(* IEC 61131-3 sources: deprecated-refusr-repo/samples (part 17) *)

(* ---- 5-MUX_stows-month-choos.st ---- *)
(*
This code implements a shuffled multiplexer with 5 control bits.
The control bits are: Data[N3], Data[N24], Data[N2], Data[N10], Data[N1]
The input bits are: Data[N22], Data[N5], Data[N4], Data[N11], Data[N6], Data[N7], Data[N21], Data[N8], Data[N9], Data[N12], Data[N20], Data[N23], Data[N17], Data[N14], Data[N25], Data[N26], Data[N28], Data[N15], Data[N30], Data[N13], Data[N16], Data[N19], Data[N27], Data[N29], Data[N18], Data[N31], Data[N34], Data[N32], Data[N33], Data[N35], Data[N36], Data[N37]

The symbolic expression is:
((((((((((((((((((((((((((((((((!(((((!(IN3)) & (!(IN24))) & (!(IN2))) & (!(IN10))) & (!(IN1)))) | IN22) & ((!((((IN3 & (!(IN24))) & (!(IN2))) & (!(IN10))) & (!(IN1)))) | IN5)) & ((!(((((!(IN3)) & IN24) & (!(IN2))) & (!(IN10))) & (!(IN1)))) | IN4)) & ((!((((IN3 & IN24) & (!(IN2))) & (!(IN10))) & (!(IN1)))) | IN11)) & ((!(((((!(IN3)) & (!(IN24))) & IN2) & (!(IN10))) & (!(IN1)))) | IN6)) & ((!((((IN3 & (!(IN24))) & IN2) & (!(IN10))) & (!(IN1)))) | IN7)) & ((!(((((!(IN3)) & IN24) & IN2) & (!(IN10))) & (!(IN1)))) | IN21)) & ((!((((IN3 & IN24) & IN2) & (!(IN10))) & (!(IN1)))) | IN8)) & ((!(((((!(IN3)) & (!(IN24))) & (!(IN2))) & IN10) & (!(IN1)))) | IN9)) & ((!((((IN3 & (!(IN24))) & (!(IN2))) & IN10) & (!(IN1)))) | IN12)) & ((!(((((!(IN3)) & IN24) & (!(IN2))) & IN10) & (!(IN1)))) | IN20)) & ((!((((IN3 & IN24) & (!(IN2))) & IN10) & (!(IN1)))) | IN23)) & ((!(((((!(IN3)) & (!(IN24))) & IN2) & IN10) & (!(IN1)))) | IN17)) & ((!((((IN3 & (!(IN24))) & IN2) & IN10) & (!(IN1)))) | IN14)) & ((!(((((!(IN3)) & IN24) & IN2) & IN10) & (!(IN1)))) | IN25)) & ((!((((IN3 & IN24) & IN2) & IN10) & (!(IN1)))) | IN26)) & ((!(((((!(IN3)) & (!(IN24))) & (!(IN2))) & (!(IN10))) & IN1)) | IN28)) & ((!((((IN3 & (!(IN24))) & (!(IN2))) & (!(IN10))) & IN1)) | IN15)) & ((!(((((!(IN3)) & IN24) & (!(IN2))) & (!(IN10))) & IN1)) | IN30)) & ((!((((IN3 & IN24) & (!(IN2))) & (!(IN10))) & IN1)) | IN13)) & ((!(((((!(IN3)) & (!(IN24))) & IN2) & (!(IN10))) & IN1)) | IN16)) & ((!((((IN3 & (!(IN24))) & IN2) & (!(IN10))) & IN1)) | IN19)) & ((!(((((!(IN3)) & IN24) & IN2) & (!(IN10))) & IN1)) | IN27)) & ((!((((IN3 & IN24) & IN2) & (!(IN10))) & IN1)) | IN29)) & ((!(((((!(IN3)) & (!(IN24))) & (!(IN2))) & IN10) & IN1)) | IN18)) & ((!((((IN3 & (!(IN24))) & (!(IN2))) & IN10) & IN1)) | IN31)) & ((!(((((!(IN3)) & IN24) & (!(IN2))) & IN10) & IN1)) | IN34)) & ((!((((IN3 & IN24) & (!(IN2))) & IN10) & IN1)) | IN32)) & ((!(((((!(IN3)) & (!(IN24))) & IN2) & IN10) & IN1)) | IN33)) & ((!((((IN3 & (!(IN24))) & IN2) & IN10) & IN1)) | IN35)) & ((!(((((!(IN3)) & IN24) & IN2) & IN10) & IN1)) | IN36)) & ((!((((IN3 & IN24) & IN2) & IN10) & IN1)) | IN37)

*)

FUNCTION_BLOCK F_CollectInput
  VAR_IN_OUT
      Data : ARRAY[1..40] OF BOOL;
  END_VAR
  VAR_INPUT
      TICK  : BOOL := 0;
      IN1   : BOOL := 0;
      IN2   : BOOL := 0;
      IN3   : BOOL := 0;
      IN4   : BOOL := 0;
      IN5   : BOOL := 0;
      RESET : BOOL := FALSE;
  END_VAR
  VAR_OUTPUT
      Finished : BOOL;
  END_VAR
  VAR
      j    : USINT := 1;
      tock : BOOL  := 0;
  END_VAR
  IF NOT RESET AND tock = NOT TICK THEN
      Data[j]   := IN1;
      Data[j+1] := IN2;
      Data[j+2] := IN3;
      Data[j+3] := IN4;
      Data[j+4] := IN5;
      j := j + 5;
      tock := TICK;
  ELSE
      j := 1;
      tock := 0;
  END_IF;
  Finished := (j > 40);
END_FUNCTION_BLOCK

PROGRAM Boiler
  VAR
    Data  : ARRAY[1..40] OF BOOL;
    Ready : BOOL;
    CollectInput : F_CollectInput;
  END_VAR
  VAR
    TICK     AT %IX1.0 : BOOL;
    IN1      AT %IX0.3 : BOOL;
    IN2      AT %IX0.4 : BOOL;
    IN3      AT %IX0.5 : BOOL;
    IN4      AT %IX0.6 : BOOL;
    IN5      AT %IX0.7 : BOOL;
    OutReady AT %QX0.0 : BOOL := FALSE;
    FeedNext AT %QX0.1 : BOOL := FALSE;
    Out      AT %QX0.2 : BOOL;
  END_VAR
  CollectInput(TICK:=TICK, IN1:=IN1, IN2:=IN2, IN3:=IN3, IN4:=IN4, IN5:=IN5);
  Ready := CollectInput.Finished;
  FeedNext := 1;
  IF Ready THEN
    Out := (((((((((((((((((((((((((((((((((NOT (((((NOT Data[3]) AND (NOT Data[24])) AND (NOT Data[2])) AND (NOT Data[10])) AND (NOT Data[1]))) OR Data[22]) AND ((NOT ((((Data[3] AND (NOT Data[24])) AND (NOT Data[2])) AND (NOT Data[10])) AND (NOT Data[1]))) OR Data[5])) AND ((NOT (((((NOT Data[3]) AND Data[24]) AND (NOT Data[2])) AND (NOT Data[10])) AND (NOT Data[1]))) OR Data[4])) AND ((NOT ((((Data[3] AND Data[24]) AND (NOT Data[2])) AND (NOT Data[10])) AND (NOT Data[1]))) OR Data[11])) AND ((NOT (((((NOT Data[3]) AND (NOT Data[24])) AND Data[2]) AND (NOT Data[10])) AND (NOT Data[1]))) OR Data[6])) AND ((NOT ((((Data[3] AND (NOT Data[24])) AND Data[2]) AND (NOT Data[10])) AND (NOT Data[1]))) OR Data[7])) AND ((NOT (((((NOT Data[3]) AND Data[24]) AND Data[2]) AND (NOT Data[10])) AND (NOT Data[1]))) OR Data[21])) AND ((NOT ((((Data[3] AND Data[24]) AND Data[2]) AND (NOT Data[10])) AND (NOT Data[1]))) OR Data[8])) AND ((NOT (((((NOT Data[3]) AND (NOT Data[24])) AND (NOT Data[2])) AND Data[10]) AND (NOT Data[1]))) OR Data[9])) AND ((NOT ((((Data[3] AND (NOT Data[24])) AND (NOT Data[2])) AND Data[10]) AND (NOT Data[1]))) OR Data[12])) AND ((NOT (((((NOT Data[3]) AND Data[24]) AND (NOT Data[2])) AND Data[10]) AND (NOT Data[1]))) OR Data[20])) AND ((NOT ((((Data[3] AND Data[24]) AND (NOT Data[2])) AND Data[10]) AND (NOT Data[1]))) OR Data[23])) AND ((NOT (((((NOT Data[3]) AND (NOT Data[24])) AND Data[2]) AND Data[10]) AND (NOT Data[1]))) OR Data[17])) AND ((NOT ((((Data[3] AND (NOT Data[24])) AND Data[2]) AND Data[10]) AND (NOT Data[1]))) OR Data[14])) AND ((NOT (((((NOT Data[3]) AND Data[24]) AND Data[2]) AND Data[10]) AND (NOT Data[1]))) OR Data[25])) AND ((NOT ((((Data[3] AND Data[24]) AND Data[2]) AND Data[10]) AND (NOT Data[1]))) OR Data[26])) AND ((NOT (((((NOT Data[3]) AND (NOT Data[24])) AND (NOT Data[2])) AND (NOT Data[10])) AND Data[1])) OR Data[28])) AND ((NOT ((((Data[3] AND (NOT Data[24])) AND (NOT Data[2])) AND (NOT Data[10])) AND Data[1])) OR Data[15])) AND ((NOT (((((NOT Data[3]) AND Data[24]) AND (NOT Data[2])) AND (NOT Data[10])) AND Data[1])) OR Data[30])) AND ((NOT ((((Data[3] AND Data[24]) AND (NOT Data[2])) AND (NOT Data[10])) AND Data[1])) OR Data[13])) AND ((NOT (((((NOT Data[3]) AND (NOT Data[24])) AND Data[2]) AND (NOT Data[10])) AND Data[1])) OR Data[16])) AND ((NOT ((((Data[3] AND (NOT Data[24])) AND Data[2]) AND (NOT Data[10])) AND Data[1])) OR Data[19])) AND ((NOT (((((NOT Data[3]) AND Data[24]) AND Data[2]) AND (NOT Data[10])) AND Data[1])) OR Data[27])) AND ((NOT ((((Data[3] AND Data[24]) AND Data[2]) AND (NOT Data[10])) AND Data[1])) OR Data[29])) AND ((NOT (((((NOT Data[3]) AND (NOT Data[24])) AND (NOT Data[2])) AND Data[10]) AND Data[1])) OR Data[18])) AND ((NOT ((((Data[3] AND (NOT Data[24])) AND (NOT Data[2])) AND Data[10]) AND Data[1])) OR Data[31])) AND ((NOT (((((NOT Data[3]) AND Data[24]) AND (NOT Data[2])) AND Data[10]) AND Data[1])) OR Data[34])) AND ((NOT ((((Data[3] AND Data[24]) AND (NOT Data[2])) AND Data[10]) AND Data[1])) OR Data[32])) AND ((NOT (((((NOT Data[3]) AND (NOT Data[24])) AND Data[2]) AND Data[10]) AND Data[1])) OR Data[33])) AND ((NOT ((((Data[3] AND (NOT Data[24])) AND Data[2]) AND Data[10]) AND Data[1])) OR Data[35])) AND ((NOT (((((NOT Data[3]) AND Data[24]) AND Data[2]) AND Data[10]) AND Data[1])) OR Data[36])) AND ((NOT ((((Data[3] AND Data[24]) AND Data[2]) AND Data[10]) AND Data[1])) OR Data[37]));
    OutReady := 1;
    CollectInput(RESET:=TRUE);
  END_IF;
END_PROGRAM

CONFIGURATION Config0
  RESOURCE Res0 ON PLC
    TASK task0(INTERVAL := T#20ms,PRIORITY := 0);
    PROGRAM instance0 WITH task0 : Boiler;
  END_RESOURCE
END_CONFIGURATION

(* ---- 5-MUX_strop-getup-abyss.st ---- *)
(*
This code implements a shuffled multiplexer with 5 control bits.
The control bits are: Data[N2], Data[N8], Data[N3], Data[N22], Data[N21]
The input bits are: Data[N20], Data[N25], Data[N5], Data[N1], Data[N6], Data[N24], Data[N23], Data[N26], Data[N27], Data[N7], Data[N28], Data[N29], Data[N10], Data[N30], Data[N33], Data[N9], Data[N4], Data[N11], Data[N12], Data[N31], Data[N32], Data[N36], Data[N34], Data[N37], Data[N15], Data[N35], Data[N14], Data[N13], Data[N17], Data[N18], Data[N16], Data[N19]

The symbolic expression is:
((((((((((((((((((((((((((((((((!(((((!(IN2)) & (!(IN8))) & (!(IN3))) & (!(IN22))) & (!(IN21)))) | IN20) & ((!((((IN2 & (!(IN8))) & (!(IN3))) & (!(IN22))) & (!(IN21)))) | IN25)) & ((!(((((!(IN2)) & IN8) & (!(IN3))) & (!(IN22))) & (!(IN21)))) | IN5)) & ((!((((IN2 & IN8) & (!(IN3))) & (!(IN22))) & (!(IN21)))) | IN1)) & ((!(((((!(IN2)) & (!(IN8))) & IN3) & (!(IN22))) & (!(IN21)))) | IN6)) & ((!((((IN2 & (!(IN8))) & IN3) & (!(IN22))) & (!(IN21)))) | IN24)) & ((!(((((!(IN2)) & IN8) & IN3) & (!(IN22))) & (!(IN21)))) | IN23)) & ((!((((IN2 & IN8) & IN3) & (!(IN22))) & (!(IN21)))) | IN26)) & ((!(((((!(IN2)) & (!(IN8))) & (!(IN3))) & IN22) & (!(IN21)))) | IN27)) & ((!((((IN2 & (!(IN8))) & (!(IN3))) & IN22) & (!(IN21)))) | IN7)) & ((!(((((!(IN2)) & IN8) & (!(IN3))) & IN22) & (!(IN21)))) | IN28)) & ((!((((IN2 & IN8) & (!(IN3))) & IN22) & (!(IN21)))) | IN29)) & ((!(((((!(IN2)) & (!(IN8))) & IN3) & IN22) & (!(IN21)))) | IN10)) & ((!((((IN2 & (!(IN8))) & IN3) & IN22) & (!(IN21)))) | IN30)) & ((!(((((!(IN2)) & IN8) & IN3) & IN22) & (!(IN21)))) | IN33)) & ((!((((IN2 & IN8) & IN3) & IN22) & (!(IN21)))) | IN9)) & ((!(((((!(IN2)) & (!(IN8))) & (!(IN3))) & (!(IN22))) & IN21)) | IN4)) & ((!((((IN2 & (!(IN8))) & (!(IN3))) & (!(IN22))) & IN21)) | IN11)) & ((!(((((!(IN2)) & IN8) & (!(IN3))) & (!(IN22))) & IN21)) | IN12)) & ((!((((IN2 & IN8) & (!(IN3))) & (!(IN22))) & IN21)) | IN31)) & ((!(((((!(IN2)) & (!(IN8))) & IN3) & (!(IN22))) & IN21)) | IN32)) & ((!((((IN2 & (!(IN8))) & IN3) & (!(IN22))) & IN21)) | IN36)) & ((!(((((!(IN2)) & IN8) & IN3) & (!(IN22))) & IN21)) | IN34)) & ((!((((IN2 & IN8) & IN3) & (!(IN22))) & IN21)) | IN37)) & ((!(((((!(IN2)) & (!(IN8))) & (!(IN3))) & IN22) & IN21)) | IN15)) & ((!((((IN2 & (!(IN8))) & (!(IN3))) & IN22) & IN21)) | IN35)) & ((!(((((!(IN2)) & IN8) & (!(IN3))) & IN22) & IN21)) | IN14)) & ((!((((IN2 & IN8) & (!(IN3))) & IN22) & IN21)) | IN13)) & ((!(((((!(IN2)) & (!(IN8))) & IN3) & IN22) & IN21)) | IN17)) & ((!((((IN2 & (!(IN8))) & IN3) & IN22) & IN21)) | IN18)) & ((!(((((!(IN2)) & IN8) & IN3) & IN22) & IN21)) | IN16)) & ((!((((IN2 & IN8) & IN3) & IN22) & IN21)) | IN19)

*)

FUNCTION_BLOCK F_CollectInput
  VAR_IN_OUT
      Data : ARRAY[1..40] OF BOOL;
  END_VAR
  VAR_INPUT
      TICK  : BOOL := 0;
      IN1   : BOOL := 0;
      IN2   : BOOL := 0;
      IN3   : BOOL := 0;
      IN4   : BOOL := 0;
      IN5   : BOOL := 0;
      RESET : BOOL := FALSE;
  END_VAR
  VAR_OUTPUT
      Finished : BOOL;
  END_VAR
  VAR
      j    : USINT := 1;
      tock : BOOL  := 0;
  END_VAR
  IF NOT RESET AND tock = NOT TICK THEN
      Data[j]   := IN1;
      Data[j+1] := IN2;
      Data[j+2] := IN3;
      Data[j+3] := IN4;
      Data[j+4] := IN5;
      j := j + 5;
      tock := TICK;
  ELSE
      j := 1;
      tock := 0;
  END_IF;
  Finished := (j > 40);
END_FUNCTION_BLOCK

PROGRAM Boiler
  VAR
    Data  : ARRAY[1..40] OF BOOL;
    Ready : BOOL;
    CollectInput : F_CollectInput;
  END_VAR
  VAR
    TICK     AT %IX1.0 : BOOL;
    IN1      AT %IX0.3 : BOOL;
    IN2      AT %IX0.4 : BOOL;
    IN3      AT %IX0.5 : BOOL;
    IN4      AT %IX0.6 : BOOL;
    IN5      AT %IX0.7 : BOOL;
    OutReady AT %QX0.0 : BOOL := FALSE;
    FeedNext AT %QX0.1 : BOOL := FALSE;
    Out      AT %QX0.2 : BOOL;
  END_VAR
  CollectInput(TICK:=TICK, IN1:=IN1, IN2:=IN2, IN3:=IN3, IN4:=IN4, IN5:=IN5);
  Ready := CollectInput.Finished;
  FeedNext := 1;
  IF Ready THEN
    Out := (((((((((((((((((((((((((((((((((NOT (((((NOT Data[2]) AND (NOT Data[8])) AND (NOT Data[3])) AND (NOT Data[22])) AND (NOT Data[21]))) OR Data[20]) AND ((NOT ((((Data[2] AND (NOT Data[8])) AND (NOT Data[3])) AND (NOT Data[22])) AND (NOT Data[21]))) OR Data[25])) AND ((NOT (((((NOT Data[2]) AND Data[8]) AND (NOT Data[3])) AND (NOT Data[22])) AND (NOT Data[21]))) OR Data[5])) AND ((NOT ((((Data[2] AND Data[8]) AND (NOT Data[3])) AND (NOT Data[22])) AND (NOT Data[21]))) OR Data[1])) AND ((NOT (((((NOT Data[2]) AND (NOT Data[8])) AND Data[3]) AND (NOT Data[22])) AND (NOT Data[21]))) OR Data[6])) AND ((NOT ((((Data[2] AND (NOT Data[8])) AND Data[3]) AND (NOT Data[22])) AND (NOT Data[21]))) OR Data[24])) AND ((NOT (((((NOT Data[2]) AND Data[8]) AND Data[3]) AND (NOT Data[22])) AND (NOT Data[21]))) OR Data[23])) AND ((NOT ((((Data[2] AND Data[8]) AND Data[3]) AND (NOT Data[22])) AND (NOT Data[21]))) OR Data[26])) AND ((NOT (((((NOT Data[2]) AND (NOT Data[8])) AND (NOT Data[3])) AND Data[22]) AND (NOT Data[21]))) OR Data[27])) AND ((NOT ((((Data[2] AND (NOT Data[8])) AND (NOT Data[3])) AND Data[22]) AND (NOT Data[21]))) OR Data[7])) AND ((NOT (((((NOT Data[2]) AND Data[8]) AND (NOT Data[3])) AND Data[22]) AND (NOT Data[21]))) OR Data[28])) AND ((NOT ((((Data[2] AND Data[8]) AND (NOT Data[3])) AND Data[22]) AND (NOT Data[21]))) OR Data[29])) AND ((NOT (((((NOT Data[2]) AND (NOT Data[8])) AND Data[3]) AND Data[22]) AND (NOT Data[21]))) OR Data[10])) AND ((NOT ((((Data[2] AND (NOT Data[8])) AND Data[3]) AND Data[22]) AND (NOT Data[21]))) OR Data[30])) AND ((NOT (((((NOT Data[2]) AND Data[8]) AND Data[3]) AND Data[22]) AND (NOT Data[21]))) OR Data[33])) AND ((NOT ((((Data[2] AND Data[8]) AND Data[3]) AND Data[22]) AND (NOT Data[21]))) OR Data[9])) AND ((NOT (((((NOT Data[2]) AND (NOT Data[8])) AND (NOT Data[3])) AND (NOT Data[22])) AND Data[21])) OR Data[4])) AND ((NOT ((((Data[2] AND (NOT Data[8])) AND (NOT Data[3])) AND (NOT Data[22])) AND Data[21])) OR Data[11])) AND ((NOT (((((NOT Data[2]) AND Data[8]) AND (NOT Data[3])) AND (NOT Data[22])) AND Data[21])) OR Data[12])) AND ((NOT ((((Data[2] AND Data[8]) AND (NOT Data[3])) AND (NOT Data[22])) AND Data[21])) OR Data[31])) AND ((NOT (((((NOT Data[2]) AND (NOT Data[8])) AND Data[3]) AND (NOT Data[22])) AND Data[21])) OR Data[32])) AND ((NOT ((((Data[2] AND (NOT Data[8])) AND Data[3]) AND (NOT Data[22])) AND Data[21])) OR Data[36])) AND ((NOT (((((NOT Data[2]) AND Data[8]) AND Data[3]) AND (NOT Data[22])) AND Data[21])) OR Data[34])) AND ((NOT ((((Data[2] AND Data[8]) AND Data[3]) AND (NOT Data[22])) AND Data[21])) OR Data[37])) AND ((NOT (((((NOT Data[2]) AND (NOT Data[8])) AND (NOT Data[3])) AND Data[22]) AND Data[21])) OR Data[15])) AND ((NOT ((((Data[2] AND (NOT Data[8])) AND (NOT Data[3])) AND Data[22]) AND Data[21])) OR Data[35])) AND ((NOT (((((NOT Data[2]) AND Data[8]) AND (NOT Data[3])) AND Data[22]) AND Data[21])) OR Data[14])) AND ((NOT ((((Data[2] AND Data[8]) AND (NOT Data[3])) AND Data[22]) AND Data[21])) OR Data[13])) AND ((NOT (((((NOT Data[2]) AND (NOT Data[8])) AND Data[3]) AND Data[22]) AND Data[21])) OR Data[17])) AND ((NOT ((((Data[2] AND (NOT Data[8])) AND Data[3]) AND Data[22]) AND Data[21])) OR Data[18])) AND ((NOT (((((NOT Data[2]) AND Data[8]) AND Data[3]) AND Data[22]) AND Data[21])) OR Data[16])) AND ((NOT ((((Data[2] AND Data[8]) AND Data[3]) AND Data[22]) AND Data[21])) OR Data[19]));
    OutReady := 1;
    CollectInput(RESET:=TRUE);
  END_IF;
END_PROGRAM

CONFIGURATION Config0
  RESOURCE Res0 ON PLC
    TASK task0(INTERVAL := T#20ms,PRIORITY := 0);
    PROGRAM instance0 WITH task0 : Boiler;
  END_RESOURCE
END_CONFIGURATION

(* ---- 5-MUX_supes-buret-rules.st ---- *)
(*
This code implements a shuffled multiplexer with 5 control bits.
The control bits are: Data[N20], Data[N2], Data[N3], Data[N1], Data[N4]
The input bits are: Data[N7], Data[N21], Data[N22], Data[N25], Data[N5], Data[N24], Data[N9], Data[N10], Data[N8], Data[N26], Data[N23], Data[N6], Data[N11], Data[N12], Data[N28], Data[N13], Data[N14], Data[N30], Data[N15], Data[N29], Data[N16], Data[N17], Data[N18], Data[N19], Data[N27], Data[N31], Data[N33], Data[N35], Data[N32], Data[N34], Data[N37], Data[N36]

The symbolic expression is:
((((((((((((((((((((((((((((((((!(((((!(IN20)) & (!(IN2))) & (!(IN3))) & (!(IN1))) & (!(IN4)))) | IN7) & ((!((((IN20 & (!(IN2))) & (!(IN3))) & (!(IN1))) & (!(IN4)))) | IN21)) & ((!(((((!(IN20)) & IN2) & (!(IN3))) & (!(IN1))) & (!(IN4)))) | IN22)) & ((!((((IN20 & IN2) & (!(IN3))) & (!(IN1))) & (!(IN4)))) | IN25)) & ((!(((((!(IN20)) & (!(IN2))) & IN3) & (!(IN1))) & (!(IN4)))) | IN5)) & ((!((((IN20 & (!(IN2))) & IN3) & (!(IN1))) & (!(IN4)))) | IN24)) & ((!(((((!(IN20)) & IN2) & IN3) & (!(IN1))) & (!(IN4)))) | IN9)) & ((!((((IN20 & IN2) & IN3) & (!(IN1))) & (!(IN4)))) | IN10)) & ((!(((((!(IN20)) & (!(IN2))) & (!(IN3))) & IN1) & (!(IN4)))) | IN8)) & ((!((((IN20 & (!(IN2))) & (!(IN3))) & IN1) & (!(IN4)))) | IN26)) & ((!(((((!(IN20)) & IN2) & (!(IN3))) & IN1) & (!(IN4)))) | IN23)) & ((!((((IN20 & IN2) & (!(IN3))) & IN1) & (!(IN4)))) | IN6)) & ((!(((((!(IN20)) & (!(IN2))) & IN3) & IN1) & (!(IN4)))) | IN11)) & ((!((((IN20 & (!(IN2))) & IN3) & IN1) & (!(IN4)))) | IN12)) & ((!(((((!(IN20)) & IN2) & IN3) & IN1) & (!(IN4)))) | IN28)) & ((!((((IN20 & IN2) & IN3) & IN1) & (!(IN4)))) | IN13)) & ((!(((((!(IN20)) & (!(IN2))) & (!(IN3))) & (!(IN1))) & IN4)) | IN14)) & ((!((((IN20 & (!(IN2))) & (!(IN3))) & (!(IN1))) & IN4)) | IN30)) & ((!(((((!(IN20)) & IN2) & (!(IN3))) & (!(IN1))) & IN4)) | IN15)) & ((!((((IN20 & IN2) & (!(IN3))) & (!(IN1))) & IN4)) | IN29)) & ((!(((((!(IN20)) & (!(IN2))) & IN3) & (!(IN1))) & IN4)) | IN16)) & ((!((((IN20 & (!(IN2))) & IN3) & (!(IN1))) & IN4)) | IN17)) & ((!(((((!(IN20)) & IN2) & IN3) & (!(IN1))) & IN4)) | IN18)) & ((!((((IN20 & IN2) & IN3) & (!(IN1))) & IN4)) | IN19)) & ((!(((((!(IN20)) & (!(IN2))) & (!(IN3))) & IN1) & IN4)) | IN27)) & ((!((((IN20 & (!(IN2))) & (!(IN3))) & IN1) & IN4)) | IN31)) & ((!(((((!(IN20)) & IN2) & (!(IN3))) & IN1) & IN4)) | IN33)) & ((!((((IN20 & IN2) & (!(IN3))) & IN1) & IN4)) | IN35)) & ((!(((((!(IN20)) & (!(IN2))) & IN3) & IN1) & IN4)) | IN32)) & ((!((((IN20 & (!(IN2))) & IN3) & IN1) & IN4)) | IN34)) & ((!(((((!(IN20)) & IN2) & IN3) & IN1) & IN4)) | IN37)) & ((!((((IN20 & IN2) & IN3) & IN1) & IN4)) | IN36)

*)

FUNCTION_BLOCK F_CollectInput
  VAR_IN_OUT
      Data : ARRAY[1..40] OF BOOL;
  END_VAR
  VAR_INPUT
      TICK  : BOOL := 0;
      IN1   : BOOL := 0;
      IN2   : BOOL := 0;
      IN3   : BOOL := 0;
      IN4   : BOOL := 0;
      IN5   : BOOL := 0;
      RESET : BOOL := FALSE;
  END_VAR
  VAR_OUTPUT
      Finished : BOOL;
  END_VAR
  VAR
      j    : USINT := 1;
      tock : BOOL  := 0;
  END_VAR
  IF NOT RESET AND tock = NOT TICK THEN
      Data[j]   := IN1;
      Data[j+1] := IN2;
      Data[j+2] := IN3;
      Data[j+3] := IN4;
      Data[j+4] := IN5;
      j := j + 5;
      tock := TICK;
  ELSE
      j := 1;
      tock := 0;
  END_IF;
  Finished := (j > 40);
END_FUNCTION_BLOCK

PROGRAM Boiler
  VAR
    Data  : ARRAY[1..40] OF BOOL;
    Ready : BOOL;
    CollectInput : F_CollectInput;
  END_VAR
  VAR
    TICK     AT %IX1.0 : BOOL;
    IN1      AT %IX0.3 : BOOL;
    IN2      AT %IX0.4 : BOOL;
    IN3      AT %IX0.5 : BOOL;
    IN4      AT %IX0.6 : BOOL;
    IN5      AT %IX0.7 : BOOL;
    OutReady AT %QX0.0 : BOOL := FALSE;
    FeedNext AT %QX0.1 : BOOL := FALSE;
    Out      AT %QX0.2 : BOOL;
  END_VAR
  CollectInput(TICK:=TICK, IN1:=IN1, IN2:=IN2, IN3:=IN3, IN4:=IN4, IN5:=IN5);
  Ready := CollectInput.Finished;
  FeedNext := 1;
  IF Ready THEN
    Out := (((((((((((((((((((((((((((((((((NOT (((((NOT Data[20]) AND (NOT Data[2])) AND (NOT Data[3])) AND (NOT Data[1])) AND (NOT Data[4]))) OR Data[7]) AND ((NOT ((((Data[20] AND (NOT Data[2])) AND (NOT Data[3])) AND (NOT Data[1])) AND (NOT Data[4]))) OR Data[21])) AND ((NOT (((((NOT Data[20]) AND Data[2]) AND (NOT Data[3])) AND (NOT Data[1])) AND (NOT Data[4]))) OR Data[22])) AND ((NOT ((((Data[20] AND Data[2]) AND (NOT Data[3])) AND (NOT Data[1])) AND (NOT Data[4]))) OR Data[25])) AND ((NOT (((((NOT Data[20]) AND (NOT Data[2])) AND Data[3]) AND (NOT Data[1])) AND (NOT Data[4]))) OR Data[5])) AND ((NOT ((((Data[20] AND (NOT Data[2])) AND Data[3]) AND (NOT Data[1])) AND (NOT Data[4]))) OR Data[24])) AND ((NOT (((((NOT Data[20]) AND Data[2]) AND Data[3]) AND (NOT Data[1])) AND (NOT Data[4]))) OR Data[9])) AND ((NOT ((((Data[20] AND Data[2]) AND Data[3]) AND (NOT Data[1])) AND (NOT Data[4]))) OR Data[10])) AND ((NOT (((((NOT Data[20]) AND (NOT Data[2])) AND (NOT Data[3])) AND Data[1]) AND (NOT Data[4]))) OR Data[8])) AND ((NOT ((((Data[20] AND (NOT Data[2])) AND (NOT Data[3])) AND Data[1]) AND (NOT Data[4]))) OR Data[26])) AND ((NOT (((((NOT Data[20]) AND Data[2]) AND (NOT Data[3])) AND Data[1]) AND (NOT Data[4]))) OR Data[23])) AND ((NOT ((((Data[20] AND Data[2]) AND (NOT Data[3])) AND Data[1]) AND (NOT Data[4]))) OR Data[6])) AND ((NOT (((((NOT Data[20]) AND (NOT Data[2])) AND Data[3]) AND Data[1]) AND (NOT Data[4]))) OR Data[11])) AND ((NOT ((((Data[20] AND (NOT Data[2])) AND Data[3]) AND Data[1]) AND (NOT Data[4]))) OR Data[12])) AND ((NOT (((((NOT Data[20]) AND Data[2]) AND Data[3]) AND Data[1]) AND (NOT Data[4]))) OR Data[28])) AND ((NOT ((((Data[20] AND Data[2]) AND Data[3]) AND Data[1]) AND (NOT Data[4]))) OR Data[13])) AND ((NOT (((((NOT Data[20]) AND (NOT Data[2])) AND (NOT Data[3])) AND (NOT Data[1])) AND Data[4])) OR Data[14])) AND ((NOT ((((Data[20] AND (NOT Data[2])) AND (NOT Data[3])) AND (NOT Data[1])) AND Data[4])) OR Data[30])) AND ((NOT (((((NOT Data[20]) AND Data[2]) AND (NOT Data[3])) AND (NOT Data[1])) AND Data[4])) OR Data[15])) AND ((NOT ((((Data[20] AND Data[2]) AND (NOT Data[3])) AND (NOT Data[1])) AND Data[4])) OR Data[29])) AND ((NOT (((((NOT Data[20]) AND (NOT Data[2])) AND Data[3]) AND (NOT Data[1])) AND Data[4])) OR Data[16])) AND ((NOT ((((Data[20] AND (NOT Data[2])) AND Data[3]) AND (NOT Data[1])) AND Data[4])) OR Data[17])) AND ((NOT (((((NOT Data[20]) AND Data[2]) AND Data[3]) AND (NOT Data[1])) AND Data[4])) OR Data[18])) AND ((NOT ((((Data[20] AND Data[2]) AND Data[3]) AND (NOT Data[1])) AND Data[4])) OR Data[19])) AND ((NOT (((((NOT Data[20]) AND (NOT Data[2])) AND (NOT Data[3])) AND Data[1]) AND Data[4])) OR Data[27])) AND ((NOT ((((Data[20] AND (NOT Data[2])) AND (NOT Data[3])) AND Data[1]) AND Data[4])) OR Data[31])) AND ((NOT (((((NOT Data[20]) AND Data[2]) AND (NOT Data[3])) AND Data[1]) AND Data[4])) OR Data[33])) AND ((NOT ((((Data[20] AND Data[2]) AND (NOT Data[3])) AND Data[1]) AND Data[4])) OR Data[35])) AND ((NOT (((((NOT Data[20]) AND (NOT Data[2])) AND Data[3]) AND Data[1]) AND Data[4])) OR Data[32])) AND ((NOT ((((Data[20] AND (NOT Data[2])) AND Data[3]) AND Data[1]) AND Data[4])) OR Data[34])) AND ((NOT (((((NOT Data[20]) AND Data[2]) AND Data[3]) AND Data[1]) AND Data[4])) OR Data[37])) AND ((NOT ((((Data[20] AND Data[2]) AND Data[3]) AND Data[1]) AND Data[4])) OR Data[36]));
    OutReady := 1;
    CollectInput(RESET:=TRUE);
  END_IF;
END_PROGRAM

CONFIGURATION Config0
  RESOURCE Res0 ON PLC
    TASK task0(INTERVAL := T#20ms,PRIORITY := 0);
    PROGRAM instance0 WITH task0 : Boiler;
  END_RESOURCE
END_CONFIGURATION

(* ---- 5-MUX_swart-booty-dozes.st ---- *)
(*
This code implements a shuffled multiplexer with 5 control bits.
The control bits are: Data[N20], Data[N21], Data[N2], Data[N1], Data[N3]
The input bits are: Data[N22], Data[N27], Data[N6], Data[N5], Data[N4], Data[N23], Data[N29], Data[N24], Data[N25], Data[N30], Data[N28], Data[N7], Data[N9], Data[N8], Data[N10], Data[N26], Data[N11], Data[N12], Data[N14], Data[N13], Data[N34], Data[N31], Data[N15], Data[N17], Data[N18], Data[N19], Data[N33], Data[N16], Data[N35], Data[N32], Data[N36], Data[N37]

The symbolic expression is:
((((((((((((((((((((((((((((((((!(((((!(IN20)) & (!(IN21))) & (!(IN2))) & (!(IN1))) & (!(IN3)))) | IN22) & ((!((((IN20 & (!(IN21))) & (!(IN2))) & (!(IN1))) & (!(IN3)))) | IN27)) & ((!(((((!(IN20)) & IN21) & (!(IN2))) & (!(IN1))) & (!(IN3)))) | IN6)) & ((!((((IN20 & IN21) & (!(IN2))) & (!(IN1))) & (!(IN3)))) | IN5)) & ((!(((((!(IN20)) & (!(IN21))) & IN2) & (!(IN1))) & (!(IN3)))) | IN4)) & ((!((((IN20 & (!(IN21))) & IN2) & (!(IN1))) & (!(IN3)))) | IN23)) & ((!(((((!(IN20)) & IN21) & IN2) & (!(IN1))) & (!(IN3)))) | IN29)) & ((!((((IN20 & IN21) & IN2) & (!(IN1))) & (!(IN3)))) | IN24)) & ((!(((((!(IN20)) & (!(IN21))) & (!(IN2))) & IN1) & (!(IN3)))) | IN25)) & ((!((((IN20 & (!(IN21))) & (!(IN2))) & IN1) & (!(IN3)))) | IN30)) & ((!(((((!(IN20)) & IN21) & (!(IN2))) & IN1) & (!(IN3)))) | IN28)) & ((!((((IN20 & IN21) & (!(IN2))) & IN1) & (!(IN3)))) | IN7)) & ((!(((((!(IN20)) & (!(IN21))) & IN2) & IN1) & (!(IN3)))) | IN9)) & ((!((((IN20 & (!(IN21))) & IN2) & IN1) & (!(IN3)))) | IN8)) & ((!(((((!(IN20)) & IN21) & IN2) & IN1) & (!(IN3)))) | IN10)) & ((!((((IN20 & IN21) & IN2) & IN1) & (!(IN3)))) | IN26)) & ((!(((((!(IN20)) & (!(IN21))) & (!(IN2))) & (!(IN1))) & IN3)) | IN11)) & ((!((((IN20 & (!(IN21))) & (!(IN2))) & (!(IN1))) & IN3)) | IN12)) & ((!(((((!(IN20)) & IN21) & (!(IN2))) & (!(IN1))) & IN3)) | IN14)) & ((!((((IN20 & IN21) & (!(IN2))) & (!(IN1))) & IN3)) | IN13)) & ((!(((((!(IN20)) & (!(IN21))) & IN2) & (!(IN1))) & IN3)) | IN34)) & ((!((((IN20 & (!(IN21))) & IN2) & (!(IN1))) & IN3)) | IN31)) & ((!(((((!(IN20)) & IN21) & IN2) & (!(IN1))) & IN3)) | IN15)) & ((!((((IN20 & IN21) & IN2) & (!(IN1))) & IN3)) | IN17)) & ((!(((((!(IN20)) & (!(IN21))) & (!(IN2))) & IN1) & IN3)) | IN18)) & ((!((((IN20 & (!(IN21))) & (!(IN2))) & IN1) & IN3)) | IN19)) & ((!(((((!(IN20)) & IN21) & (!(IN2))) & IN1) & IN3)) | IN33)) & ((!((((IN20 & IN21) & (!(IN2))) & IN1) & IN3)) | IN16)) & ((!(((((!(IN20)) & (!(IN21))) & IN2) & IN1) & IN3)) | IN35)) & ((!((((IN20 & (!(IN21))) & IN2) & IN1) & IN3)) | IN32)) & ((!(((((!(IN20)) & IN21) & IN2) & IN1) & IN3)) | IN36)) & ((!((((IN20 & IN21) & IN2) & IN1) & IN3)) | IN37)

*)

FUNCTION_BLOCK F_CollectInput
  VAR_IN_OUT
      Data : ARRAY[1..40] OF BOOL;
  END_VAR
  VAR_INPUT
      TICK  : BOOL := 0;
      IN1   : BOOL := 0;
      IN2   : BOOL := 0;
      IN3   : BOOL := 0;
      IN4   : BOOL := 0;
      IN5   : BOOL := 0;
      RESET : BOOL := FALSE;
  END_VAR
  VAR_OUTPUT
      Finished : BOOL;
  END_VAR
  VAR
      j    : USINT := 1;
      tock : BOOL  := 0;
  END_VAR
  IF NOT RESET AND tock = NOT TICK THEN
      Data[j]   := IN1;
      Data[j+1] := IN2;
      Data[j+2] := IN3;
      Data[j+3] := IN4;
      Data[j+4] := IN5;
      j := j + 5;
      tock := TICK;
  ELSE
      j := 1;
      tock := 0;
  END_IF;
  Finished := (j > 40);
END_FUNCTION_BLOCK

PROGRAM Boiler
  VAR
    Data  : ARRAY[1..40] OF BOOL;
    Ready : BOOL;
    CollectInput : F_CollectInput;
  END_VAR
  VAR
    TICK     AT %IX1.0 : BOOL;
    IN1      AT %IX0.3 : BOOL;
    IN2      AT %IX0.4 : BOOL;
    IN3      AT %IX0.5 : BOOL;
    IN4      AT %IX0.6 : BOOL;
    IN5      AT %IX0.7 : BOOL;
    OutReady AT %QX0.0 : BOOL := FALSE;
    FeedNext AT %QX0.1 : BOOL := FALSE;
    Out      AT %QX0.2 : BOOL;
  END_VAR
  CollectInput(TICK:=TICK, IN1:=IN1, IN2:=IN2, IN3:=IN3, IN4:=IN4, IN5:=IN5);
  Ready := CollectInput.Finished;
  FeedNext := 1;
  IF Ready THEN
    Out := (((((((((((((((((((((((((((((((((NOT (((((NOT Data[20]) AND (NOT Data[21])) AND (NOT Data[2])) AND (NOT Data[1])) AND (NOT Data[3]))) OR Data[22]) AND ((NOT ((((Data[20] AND (NOT Data[21])) AND (NOT Data[2])) AND (NOT Data[1])) AND (NOT Data[3]))) OR Data[27])) AND ((NOT (((((NOT Data[20]) AND Data[21]) AND (NOT Data[2])) AND (NOT Data[1])) AND (NOT Data[3]))) OR Data[6])) AND ((NOT ((((Data[20] AND Data[21]) AND (NOT Data[2])) AND (NOT Data[1])) AND (NOT Data[3]))) OR Data[5])) AND ((NOT (((((NOT Data[20]) AND (NOT Data[21])) AND Data[2]) AND (NOT Data[1])) AND (NOT Data[3]))) OR Data[4])) AND ((NOT ((((Data[20] AND (NOT Data[21])) AND Data[2]) AND (NOT Data[1])) AND (NOT Data[3]))) OR Data[23])) AND ((NOT (((((NOT Data[20]) AND Data[21]) AND Data[2]) AND (NOT Data[1])) AND (NOT Data[3]))) OR Data[29])) AND ((NOT ((((Data[20] AND Data[21]) AND Data[2]) AND (NOT Data[1])) AND (NOT Data[3]))) OR Data[24])) AND ((NOT (((((NOT Data[20]) AND (NOT Data[21])) AND (NOT Data[2])) AND Data[1]) AND (NOT Data[3]))) OR Data[25])) AND ((NOT ((((Data[20] AND (NOT Data[21])) AND (NOT Data[2])) AND Data[1]) AND (NOT Data[3]))) OR Data[30])) AND ((NOT (((((NOT Data[20]) AND Data[21]) AND (NOT Data[2])) AND Data[1]) AND (NOT Data[3]))) OR Data[28])) AND ((NOT ((((Data[20] AND Data[21]) AND (NOT Data[2])) AND Data[1]) AND (NOT Data[3]))) OR Data[7])) AND ((NOT (((((NOT Data[20]) AND (NOT Data[21])) AND Data[2]) AND Data[1]) AND (NOT Data[3]))) OR Data[9])) AND ((NOT ((((Data[20] AND (NOT Data[21])) AND Data[2]) AND Data[1]) AND (NOT Data[3]))) OR Data[8])) AND ((NOT (((((NOT Data[20]) AND Data[21]) AND Data[2]) AND Data[1]) AND (NOT Data[3]))) OR Data[10])) AND ((NOT ((((Data[20] AND Data[21]) AND Data[2]) AND Data[1]) AND (NOT Data[3]))) OR Data[26])) AND ((NOT (((((NOT Data[20]) AND (NOT Data[21])) AND (NOT Data[2])) AND (NOT Data[1])) AND Data[3])) OR Data[11])) AND ((NOT ((((Data[20] AND (NOT Data[21])) AND (NOT Data[2])) AND (NOT Data[1])) AND Data[3])) OR Data[12])) AND ((NOT (((((NOT Data[20]) AND Data[21]) AND (NOT Data[2])) AND (NOT Data[1])) AND Data[3])) OR Data[14])) AND ((NOT ((((Data[20] AND Data[21]) AND (NOT Data[2])) AND (NOT Data[1])) AND Data[3])) OR Data[13])) AND ((NOT (((((NOT Data[20]) AND (NOT Data[21])) AND Data[2]) AND (NOT Data[1])) AND Data[3])) OR Data[34])) AND ((NOT ((((Data[20] AND (NOT Data[21])) AND Data[2]) AND (NOT Data[1])) AND Data[3])) OR Data[31])) AND ((NOT (((((NOT Data[20]) AND Data[21]) AND Data[2]) AND (NOT Data[1])) AND Data[3])) OR Data[15])) AND ((NOT ((((Data[20] AND Data[21]) AND Data[2]) AND (NOT Data[1])) AND Data[3])) OR Data[17])) AND ((NOT (((((NOT Data[20]) AND (NOT Data[21])) AND (NOT Data[2])) AND Data[1]) AND Data[3])) OR Data[18])) AND ((NOT ((((Data[20] AND (NOT Data[21])) AND (NOT Data[2])) AND Data[1]) AND Data[3])) OR Data[19])) AND ((NOT (((((NOT Data[20]) AND Data[21]) AND (NOT Data[2])) AND Data[1]) AND Data[3])) OR Data[33])) AND ((NOT ((((Data[20] AND Data[21]) AND (NOT Data[2])) AND Data[1]) AND Data[3])) OR Data[16])) AND ((NOT (((((NOT Data[20]) AND (NOT Data[21])) AND Data[2]) AND Data[1]) AND Data[3])) OR Data[35])) AND ((NOT ((((Data[20] AND (NOT Data[21])) AND Data[2]) AND Data[1]) AND Data[3])) OR Data[32])) AND ((NOT (((((NOT Data[20]) AND Data[21]) AND Data[2]) AND Data[1]) AND Data[3])) OR Data[36])) AND ((NOT ((((Data[20] AND Data[21]) AND Data[2]) AND Data[1]) AND Data[3])) OR Data[37]));
    OutReady := 1;
    CollectInput(RESET:=TRUE);
  END_IF;
END_PROGRAM

CONFIGURATION Config0
  RESOURCE Res0 ON PLC
    TASK task0(INTERVAL := T#20ms,PRIORITY := 0);
    PROGRAM instance0 WITH task0 : Boiler;
  END_RESOURCE
END_CONFIGURATION

(* ---- 5-MUX_tamps-cluck-liras.st ---- *)
(*
This code implements a shuffled multiplexer with 5 control bits.
The control bits are: Data[N26], Data[N21], Data[N20], Data[N2], Data[N22]
The input bits are: Data[N3], Data[N1], Data[N23], Data[N24], Data[N5], Data[N4], Data[N25], Data[N6], Data[N8], Data[N10], Data[N28], Data[N27], Data[N32], Data[N11], Data[N7], Data[N29], Data[N13], Data[N15], Data[N9], Data[N14], Data[N30], Data[N31], Data[N12], Data[N16], Data[N19], Data[N17], Data[N18], Data[N34], Data[N33], Data[N36], Data[N37], Data[N35]

The symbolic expression is:
((((((((((((((((((((((((((((((((!(((((!(IN26)) & (!(IN21))) & (!(IN20))) & (!(IN2))) & (!(IN22)))) | IN3) & ((!((((IN26 & (!(IN21))) & (!(IN20))) & (!(IN2))) & (!(IN22)))) | IN1)) & ((!(((((!(IN26)) & IN21) & (!(IN20))) & (!(IN2))) & (!(IN22)))) | IN23)) & ((!((((IN26 & IN21) & (!(IN20))) & (!(IN2))) & (!(IN22)))) | IN24)) & ((!(((((!(IN26)) & (!(IN21))) & IN20) & (!(IN2))) & (!(IN22)))) | IN5)) & ((!((((IN26 & (!(IN21))) & IN20) & (!(IN2))) & (!(IN22)))) | IN4)) & ((!(((((!(IN26)) & IN21) & IN20) & (!(IN2))) & (!(IN22)))) | IN25)) & ((!((((IN26 & IN21) & IN20) & (!(IN2))) & (!(IN22)))) | IN6)) & ((!(((((!(IN26)) & (!(IN21))) & (!(IN20))) & IN2) & (!(IN22)))) | IN8)) & ((!((((IN26 & (!(IN21))) & (!(IN20))) & IN2) & (!(IN22)))) | IN10)) & ((!(((((!(IN26)) & IN21) & (!(IN20))) & IN2) & (!(IN22)))) | IN28)) & ((!((((IN26 & IN21) & (!(IN20))) & IN2) & (!(IN22)))) | IN27)) & ((!(((((!(IN26)) & (!(IN21))) & IN20) & IN2) & (!(IN22)))) | IN32)) & ((!((((IN26 & (!(IN21))) & IN20) & IN2) & (!(IN22)))) | IN11)) & ((!(((((!(IN26)) & IN21) & IN20) & IN2) & (!(IN22)))) | IN7)) & ((!((((IN26 & IN21) & IN20) & IN2) & (!(IN22)))) | IN29)) & ((!(((((!(IN26)) & (!(IN21))) & (!(IN20))) & (!(IN2))) & IN22)) | IN13)) & ((!((((IN26 & (!(IN21))) & (!(IN20))) & (!(IN2))) & IN22)) | IN15)) & ((!(((((!(IN26)) & IN21) & (!(IN20))) & (!(IN2))) & IN22)) | IN9)) & ((!((((IN26 & IN21) & (!(IN20))) & (!(IN2))) & IN22)) | IN14)) & ((!(((((!(IN26)) & (!(IN21))) & IN20) & (!(IN2))) & IN22)) | IN30)) & ((!((((IN26 & (!(IN21))) & IN20) & (!(IN2))) & IN22)) | IN31)) & ((!(((((!(IN26)) & IN21) & IN20) & (!(IN2))) & IN22)) | IN12)) & ((!((((IN26 & IN21) & IN20) & (!(IN2))) & IN22)) | IN16)) & ((!(((((!(IN26)) & (!(IN21))) & (!(IN20))) & IN2) & IN22)) | IN19)) & ((!((((IN26 & (!(IN21))) & (!(IN20))) & IN2) & IN22)) | IN17)) & ((!(((((!(IN26)) & IN21) & (!(IN20))) & IN2) & IN22)) | IN18)) & ((!((((IN26 & IN21) & (!(IN20))) & IN2) & IN22)) | IN34)) & ((!(((((!(IN26)) & (!(IN21))) & IN20) & IN2) & IN22)) | IN33)) & ((!((((IN26 & (!(IN21))) & IN20) & IN2) & IN22)) | IN36)) & ((!(((((!(IN26)) & IN21) & IN20) & IN2) & IN22)) | IN37)) & ((!((((IN26 & IN21) & IN20) & IN2) & IN22)) | IN35)

*)

FUNCTION_BLOCK F_CollectInput
  VAR_IN_OUT
      Data : ARRAY[1..40] OF BOOL;
  END_VAR
  VAR_INPUT
      TICK  : BOOL := 0;
      IN1   : BOOL := 0;
      IN2   : BOOL := 0;
      IN3   : BOOL := 0;
      IN4   : BOOL := 0;
      IN5   : BOOL := 0;
      RESET : BOOL := FALSE;
  END_VAR
  VAR_OUTPUT
      Finished : BOOL;
  END_VAR
  VAR
      j    : USINT := 1;
      tock : BOOL  := 0;
  END_VAR
  IF NOT RESET AND tock = NOT TICK THEN
      Data[j]   := IN1;
      Data[j+1] := IN2;
      Data[j+2] := IN3;
      Data[j+3] := IN4;
      Data[j+4] := IN5;
      j := j + 5;
      tock := TICK;
  ELSE
      j := 1;
      tock := 0;
  END_IF;
  Finished := (j > 40);
END_FUNCTION_BLOCK

PROGRAM Boiler
  VAR
    Data  : ARRAY[1..40] OF BOOL;
    Ready : BOOL;
    CollectInput : F_CollectInput;
  END_VAR
  VAR
    TICK     AT %IX1.0 : BOOL;
    IN1      AT %IX0.3 : BOOL;
    IN2      AT %IX0.4 : BOOL;
    IN3      AT %IX0.5 : BOOL;
    IN4      AT %IX0.6 : BOOL;
    IN5      AT %IX0.7 : BOOL;
    OutReady AT %QX0.0 : BOOL := FALSE;
    FeedNext AT %QX0.1 : BOOL := FALSE;
    Out      AT %QX0.2 : BOOL;
  END_VAR
  CollectInput(TICK:=TICK, IN1:=IN1, IN2:=IN2, IN3:=IN3, IN4:=IN4, IN5:=IN5);
  Ready := CollectInput.Finished;
  FeedNext := 1;
  IF Ready THEN
    Out := (((((((((((((((((((((((((((((((((NOT (((((NOT Data[26]) AND (NOT Data[21])) AND (NOT Data[20])) AND (NOT Data[2])) AND (NOT Data[22]))) OR Data[3]) AND ((NOT ((((Data[26] AND (NOT Data[21])) AND (NOT Data[20])) AND (NOT Data[2])) AND (NOT Data[22]))) OR Data[1])) AND ((NOT (((((NOT Data[26]) AND Data[21]) AND (NOT Data[20])) AND (NOT Data[2])) AND (NOT Data[22]))) OR Data[23])) AND ((NOT ((((Data[26] AND Data[21]) AND (NOT Data[20])) AND (NOT Data[2])) AND (NOT Data[22]))) OR Data[24])) AND ((NOT (((((NOT Data[26]) AND (NOT Data[21])) AND Data[20]) AND (NOT Data[2])) AND (NOT Data[22]))) OR Data[5])) AND ((NOT ((((Data[26] AND (NOT Data[21])) AND Data[20]) AND (NOT Data[2])) AND (NOT Data[22]))) OR Data[4])) AND ((NOT (((((NOT Data[26]) AND Data[21]) AND Data[20]) AND (NOT Data[2])) AND (NOT Data[22]))) OR Data[25])) AND ((NOT ((((Data[26] AND Data[21]) AND Data[20]) AND (NOT Data[2])) AND (NOT Data[22]))) OR Data[6])) AND ((NOT (((((NOT Data[26]) AND (NOT Data[21])) AND (NOT Data[20])) AND Data[2]) AND (NOT Data[22]))) OR Data[8])) AND ((NOT ((((Data[26] AND (NOT Data[21])) AND (NOT Data[20])) AND Data[2]) AND (NOT Data[22]))) OR Data[10])) AND ((NOT (((((NOT Data[26]) AND Data[21]) AND (NOT Data[20])) AND Data[2]) AND (NOT Data[22]))) OR Data[28])) AND ((NOT ((((Data[26] AND Data[21]) AND (NOT Data[20])) AND Data[2]) AND (NOT Data[22]))) OR Data[27])) AND ((NOT (((((NOT Data[26]) AND (NOT Data[21])) AND Data[20]) AND Data[2]) AND (NOT Data[22]))) OR Data[32])) AND ((NOT ((((Data[26] AND (NOT Data[21])) AND Data[20]) AND Data[2]) AND (NOT Data[22]))) OR Data[11])) AND ((NOT (((((NOT Data[26]) AND Data[21]) AND Data[20]) AND Data[2]) AND (NOT Data[22]))) OR Data[7])) AND ((NOT ((((Data[26] AND Data[21]) AND Data[20]) AND Data[2]) AND (NOT Data[22]))) OR Data[29])) AND ((NOT (((((NOT Data[26]) AND (NOT Data[21])) AND (NOT Data[20])) AND (NOT Data[2])) AND Data[22])) OR Data[13])) AND ((NOT ((((Data[26] AND (NOT Data[21])) AND (NOT Data[20])) AND (NOT Data[2])) AND Data[22])) OR Data[15])) AND ((NOT (((((NOT Data[26]) AND Data[21]) AND (NOT Data[20])) AND (NOT Data[2])) AND Data[22])) OR Data[9])) AND ((NOT ((((Data[26] AND Data[21]) AND (NOT Data[20])) AND (NOT Data[2])) AND Data[22])) OR Data[14])) AND ((NOT (((((NOT Data[26]) AND (NOT Data[21])) AND Data[20]) AND (NOT Data[2])) AND Data[22])) OR Data[30])) AND ((NOT ((((Data[26] AND (NOT Data[21])) AND Data[20]) AND (NOT Data[2])) AND Data[22])) OR Data[31])) AND ((NOT (((((NOT Data[26]) AND Data[21]) AND Data[20]) AND (NOT Data[2])) AND Data[22])) OR Data[12])) AND ((NOT ((((Data[26] AND Data[21]) AND Data[20]) AND (NOT Data[2])) AND Data[22])) OR Data[16])) AND ((NOT (((((NOT Data[26]) AND (NOT Data[21])) AND (NOT Data[20])) AND Data[2]) AND Data[22])) OR Data[19])) AND ((NOT ((((Data[26] AND (NOT Data[21])) AND (NOT Data[20])) AND Data[2]) AND Data[22])) OR Data[17])) AND ((NOT (((((NOT Data[26]) AND Data[21]) AND (NOT Data[20])) AND Data[2]) AND Data[22])) OR Data[18])) AND ((NOT ((((Data[26] AND Data[21]) AND (NOT Data[20])) AND Data[2]) AND Data[22])) OR Data[34])) AND ((NOT (((((NOT Data[26]) AND (NOT Data[21])) AND Data[20]) AND Data[2]) AND Data[22])) OR Data[33])) AND ((NOT ((((Data[26] AND (NOT Data[21])) AND Data[20]) AND Data[2]) AND Data[22])) OR Data[36])) AND ((NOT (((((NOT Data[26]) AND Data[21]) AND Data[20]) AND Data[2]) AND Data[22])) OR Data[37])) AND ((NOT ((((Data[26] AND Data[21]) AND Data[20]) AND Data[2]) AND Data[22])) OR Data[35]));
    OutReady := 1;
    CollectInput(RESET:=TRUE);
  END_IF;
END_PROGRAM

CONFIGURATION Config0
  RESOURCE Res0 ON PLC
    TASK task0(INTERVAL := T#20ms,PRIORITY := 0);
    PROGRAM instance0 WITH task0 : Boiler;
  END_RESOURCE
END_CONFIGURATION

(* ---- 5-MUX_tarns-bueno-oaths.st ---- *)
(*
This code implements a shuffled multiplexer with 5 control bits.
The control bits are: Data[N20], Data[N21], Data[N24], Data[N2], Data[N1]
The input bits are: Data[N25], Data[N3], Data[N7], Data[N4], Data[N6], Data[N8], Data[N5], Data[N22], Data[N23], Data[N10], Data[N26], Data[N27], Data[N28], Data[N30], Data[N9], Data[N11], Data[N12], Data[N13], Data[N29], Data[N17], Data[N14], Data[N15], Data[N16], Data[N18], Data[N31], Data[N35], Data[N19], Data[N33], Data[N32], Data[N37], Data[N36], Data[N34]

The symbolic expression is:
((((((((((((((((((((((((((((((((!(((((!(IN20)) & (!(IN21))) & (!(IN24))) & (!(IN2))) & (!(IN1)))) | IN25) & ((!((((IN20 & (!(IN21))) & (!(IN24))) & (!(IN2))) & (!(IN1)))) | IN3)) & ((!(((((!(IN20)) & IN21) & (!(IN24))) & (!(IN2))) & (!(IN1)))) | IN7)) & ((!((((IN20 & IN21) & (!(IN24))) & (!(IN2))) & (!(IN1)))) | IN4)) & ((!(((((!(IN20)) & (!(IN21))) & IN24) & (!(IN2))) & (!(IN1)))) | IN6)) & ((!((((IN20 & (!(IN21))) & IN24) & (!(IN2))) & (!(IN1)))) | IN8)) & ((!(((((!(IN20)) & IN21) & IN24) & (!(IN2))) & (!(IN1)))) | IN5)) & ((!((((IN20 & IN21) & IN24) & (!(IN2))) & (!(IN1)))) | IN22)) & ((!(((((!(IN20)) & (!(IN21))) & (!(IN24))) & IN2) & (!(IN1)))) | IN23)) & ((!((((IN20 & (!(IN21))) & (!(IN24))) & IN2) & (!(IN1)))) | IN10)) & ((!(((((!(IN20)) & IN21) & (!(IN24))) & IN2) & (!(IN1)))) | IN26)) & ((!((((IN20 & IN21) & (!(IN24))) & IN2) & (!(IN1)))) | IN27)) & ((!(((((!(IN20)) & (!(IN21))) & IN24) & IN2) & (!(IN1)))) | IN28)) & ((!((((IN20 & (!(IN21))) & IN24) & IN2) & (!(IN1)))) | IN30)) & ((!(((((!(IN20)) & IN21) & IN24) & IN2) & (!(IN1)))) | IN9)) & ((!((((IN20 & IN21) & IN24) & IN2) & (!(IN1)))) | IN11)) & ((!(((((!(IN20)) & (!(IN21))) & (!(IN24))) & (!(IN2))) & IN1)) | IN12)) & ((!((((IN20 & (!(IN21))) & (!(IN24))) & (!(IN2))) & IN1)) | IN13)) & ((!(((((!(IN20)) & IN21) & (!(IN24))) & (!(IN2))) & IN1)) | IN29)) & ((!((((IN20 & IN21) & (!(IN24))) & (!(IN2))) & IN1)) | IN17)) & ((!(((((!(IN20)) & (!(IN21))) & IN24) & (!(IN2))) & IN1)) | IN14)) & ((!((((IN20 & (!(IN21))) & IN24) & (!(IN2))) & IN1)) | IN15)) & ((!(((((!(IN20)) & IN21) & IN24) & (!(IN2))) & IN1)) | IN16)) & ((!((((IN20 & IN21) & IN24) & (!(IN2))) & IN1)) | IN18)) & ((!(((((!(IN20)) & (!(IN21))) & (!(IN24))) & IN2) & IN1)) | IN31)) & ((!((((IN20 & (!(IN21))) & (!(IN24))) & IN2) & IN1)) | IN35)) & ((!(((((!(IN20)) & IN21) & (!(IN24))) & IN2) & IN1)) | IN19)) & ((!((((IN20 & IN21) & (!(IN24))) & IN2) & IN1)) | IN33)) & ((!(((((!(IN20)) & (!(IN21))) & IN24) & IN2) & IN1)) | IN32)) & ((!((((IN20 & (!(IN21))) & IN24) & IN2) & IN1)) | IN37)) & ((!(((((!(IN20)) & IN21) & IN24) & IN2) & IN1)) | IN36)) & ((!((((IN20 & IN21) & IN24) & IN2) & IN1)) | IN34)

*)

FUNCTION_BLOCK F_CollectInput
  VAR_IN_OUT
      Data : ARRAY[1..40] OF BOOL;
  END_VAR
  VAR_INPUT
      TICK  : BOOL := 0;
      IN1   : BOOL := 0;
      IN2   : BOOL := 0;
      IN3   : BOOL := 0;
      IN4   : BOOL := 0;
      IN5   : BOOL := 0;
      RESET : BOOL := FALSE;
  END_VAR
  VAR_OUTPUT
      Finished : BOOL;
  END_VAR
  VAR
      j    : USINT := 1;
      tock : BOOL  := 0;
  END_VAR
  IF NOT RESET AND tock = NOT TICK THEN
      Data[j]   := IN1;
      Data[j+1] := IN2;
      Data[j+2] := IN3;
      Data[j+3] := IN4;
      Data[j+4] := IN5;
      j := j + 5;
      tock := TICK;
  ELSE
      j := 1;
      tock := 0;
  END_IF;
  Finished := (j > 40);
END_FUNCTION_BLOCK

PROGRAM Boiler
  VAR
    Data  : ARRAY[1..40] OF BOOL;
    Ready : BOOL;
    CollectInput : F_CollectInput;
  END_VAR
  VAR
    TICK     AT %IX1.0 : BOOL;
    IN1      AT %IX0.3 : BOOL;
    IN2      AT %IX0.4 : BOOL;
    IN3      AT %IX0.5 : BOOL;
    IN4      AT %IX0.6 : BOOL;
    IN5      AT %IX0.7 : BOOL;
    OutReady AT %QX0.0 : BOOL := FALSE;
    FeedNext AT %QX0.1 : BOOL := FALSE;
    Out      AT %QX0.2 : BOOL;
  END_VAR
  CollectInput(TICK:=TICK, IN1:=IN1, IN2:=IN2, IN3:=IN3, IN4:=IN4, IN5:=IN5);
  Ready := CollectInput.Finished;
  FeedNext := 1;
  IF Ready THEN
    Out := (((((((((((((((((((((((((((((((((NOT (((((NOT Data[20]) AND (NOT Data[21])) AND (NOT Data[24])) AND (NOT Data[2])) AND (NOT Data[1]))) OR Data[25]) AND ((NOT ((((Data[20] AND (NOT Data[21])) AND (NOT Data[24])) AND (NOT Data[2])) AND (NOT Data[1]))) OR Data[3])) AND ((NOT (((((NOT Data[20]) AND Data[21]) AND (NOT Data[24])) AND (NOT Data[2])) AND (NOT Data[1]))) OR Data[7])) AND ((NOT ((((Data[20] AND Data[21]) AND (NOT Data[24])) AND (NOT Data[2])) AND (NOT Data[1]))) OR Data[4])) AND ((NOT (((((NOT Data[20]) AND (NOT Data[21])) AND Data[24]) AND (NOT Data[2])) AND (NOT Data[1]))) OR Data[6])) AND ((NOT ((((Data[20] AND (NOT Data[21])) AND Data[24]) AND (NOT Data[2])) AND (NOT Data[1]))) OR Data[8])) AND ((NOT (((((NOT Data[20]) AND Data[21]) AND Data[24]) AND (NOT Data[2])) AND (NOT Data[1]))) OR Data[5])) AND ((NOT ((((Data[20] AND Data[21]) AND Data[24]) AND (NOT Data[2])) AND (NOT Data[1]))) OR Data[22])) AND ((NOT (((((NOT Data[20]) AND (NOT Data[21])) AND (NOT Data[24])) AND Data[2]) AND (NOT Data[1]))) OR Data[23])) AND ((NOT ((((Data[20] AND (NOT Data[21])) AND (NOT Data[24])) AND Data[2]) AND (NOT Data[1]))) OR Data[10])) AND ((NOT (((((NOT Data[20]) AND Data[21]) AND (NOT Data[24])) AND Data[2]) AND (NOT Data[1]))) OR Data[26])) AND ((NOT ((((Data[20] AND Data[21]) AND (NOT Data[24])) AND Data[2]) AND (NOT Data[1]))) OR Data[27])) AND ((NOT (((((NOT Data[20]) AND (NOT Data[21])) AND Data[24]) AND Data[2]) AND (NOT Data[1]))) OR Data[28])) AND ((NOT ((((Data[20] AND (NOT Data[21])) AND Data[24]) AND Data[2]) AND (NOT Data[1]))) OR Data[30])) AND ((NOT (((((NOT Data[20]) AND Data[21]) AND Data[24]) AND Data[2]) AND (NOT Data[1]))) OR Data[9])) AND ((NOT ((((Data[20] AND Data[21]) AND Data[24]) AND Data[2]) AND (NOT Data[1]))) OR Data[11])) AND ((NOT (((((NOT Data[20]) AND (NOT Data[21])) AND (NOT Data[24])) AND (NOT Data[2])) AND Data[1])) OR Data[12])) AND ((NOT ((((Data[20] AND (NOT Data[21])) AND (NOT Data[24])) AND (NOT Data[2])) AND Data[1])) OR Data[13])) AND ((NOT (((((NOT Data[20]) AND Data[21]) AND (NOT Data[24])) AND (NOT Data[2])) AND Data[1])) OR Data[29])) AND ((NOT ((((Data[20] AND Data[21]) AND (NOT Data[24])) AND (NOT Data[2])) AND Data[1])) OR Data[17])) AND ((NOT (((((NOT Data[20]) AND (NOT Data[21])) AND Data[24]) AND (NOT Data[2])) AND Data[1])) OR Data[14])) AND ((NOT ((((Data[20] AND (NOT Data[21])) AND Data[24]) AND (NOT Data[2])) AND Data[1])) OR Data[15])) AND ((NOT (((((NOT Data[20]) AND Data[21]) AND Data[24]) AND (NOT Data[2])) AND Data[1])) OR Data[16])) AND ((NOT ((((Data[20] AND Data[21]) AND Data[24]) AND (NOT Data[2])) AND Data[1])) OR Data[18])) AND ((NOT (((((NOT Data[20]) AND (NOT Data[21])) AND (NOT Data[24])) AND Data[2]) AND Data[1])) OR Data[31])) AND ((NOT ((((Data[20] AND (NOT Data[21])) AND (NOT Data[24])) AND Data[2]) AND Data[1])) OR Data[35])) AND ((NOT (((((NOT Data[20]) AND Data[21]) AND (NOT Data[24])) AND Data[2]) AND Data[1])) OR Data[19])) AND ((NOT ((((Data[20] AND Data[21]) AND (NOT Data[24])) AND Data[2]) AND Data[1])) OR Data[33])) AND ((NOT (((((NOT Data[20]) AND (NOT Data[21])) AND Data[24]) AND Data[2]) AND Data[1])) OR Data[32])) AND ((NOT ((((Data[20] AND (NOT Data[21])) AND Data[24]) AND Data[2]) AND Data[1])) OR Data[37])) AND ((NOT (((((NOT Data[20]) AND Data[21]) AND Data[24]) AND Data[2]) AND Data[1])) OR Data[36])) AND ((NOT ((((Data[20] AND Data[21]) AND Data[24]) AND Data[2]) AND Data[1])) OR Data[34]));
    OutReady := 1;
    CollectInput(RESET:=TRUE);
  END_IF;
END_PROGRAM

CONFIGURATION Config0
  RESOURCE Res0 ON PLC
    TASK task0(INTERVAL := T#20ms,PRIORITY := 0);
    PROGRAM instance0 WITH task0 : Boiler;
  END_RESOURCE
END_CONFIGURATION

(* ---- 5-MUX_techy-cavil-twiny.st ---- *)
(*
This code implements a shuffled multiplexer with 5 control bits.
The control bits are: Data[N21], Data[N2], Data[N1], Data[N20], Data[N22]
The input bits are: Data[N3], Data[N24], Data[N23], Data[N25], Data[N28], Data[N6], Data[N4], Data[N26], Data[N29], Data[N30], Data[N7], Data[N8], Data[N34], Data[N5], Data[N16], Data[N17], Data[N10], Data[N32], Data[N33], Data[N15], Data[N12], Data[N11], Data[N9], Data[N13], Data[N27], Data[N14], Data[N31], Data[N35], Data[N36], Data[N18], Data[N19], Data[N37]

The symbolic expression is:
((((((((((((((((((((((((((((((((!(((((!(IN21)) & (!(IN2))) & (!(IN1))) & (!(IN20))) & (!(IN22)))) | IN3) & ((!((((IN21 & (!(IN2))) & (!(IN1))) & (!(IN20))) & (!(IN22)))) | IN24)) & ((!(((((!(IN21)) & IN2) & (!(IN1))) & (!(IN20))) & (!(IN22)))) | IN23)) & ((!((((IN21 & IN2) & (!(IN1))) & (!(IN20))) & (!(IN22)))) | IN25)) & ((!(((((!(IN21)) & (!(IN2))) & IN1) & (!(IN20))) & (!(IN22)))) | IN28)) & ((!((((IN21 & (!(IN2))) & IN1) & (!(IN20))) & (!(IN22)))) | IN6)) & ((!(((((!(IN21)) & IN2) & IN1) & (!(IN20))) & (!(IN22)))) | IN4)) & ((!((((IN21 & IN2) & IN1) & (!(IN20))) & (!(IN22)))) | IN26)) & ((!(((((!(IN21)) & (!(IN2))) & (!(IN1))) & IN20) & (!(IN22)))) | IN29)) & ((!((((IN21 & (!(IN2))) & (!(IN1))) & IN20) & (!(IN22)))) | IN30)) & ((!(((((!(IN21)) & IN2) & (!(IN1))) & IN20) & (!(IN22)))) | IN7)) & ((!((((IN21 & IN2) & (!(IN1))) & IN20) & (!(IN22)))) | IN8)) & ((!(((((!(IN21)) & (!(IN2))) & IN1) & IN20) & (!(IN22)))) | IN34)) & ((!((((IN21 & (!(IN2))) & IN1) & IN20) & (!(IN22)))) | IN5)) & ((!(((((!(IN21)) & IN2) & IN1) & IN20) & (!(IN22)))) | IN16)) & ((!((((IN21 & IN2) & IN1) & IN20) & (!(IN22)))) | IN17)) & ((!(((((!(IN21)) & (!(IN2))) & (!(IN1))) & (!(IN20))) & IN22)) | IN10)) & ((!((((IN21 & (!(IN2))) & (!(IN1))) & (!(IN20))) & IN22)) | IN32)) & ((!(((((!(IN21)) & IN2) & (!(IN1))) & (!(IN20))) & IN22)) | IN33)) & ((!((((IN21 & IN2) & (!(IN1))) & (!(IN20))) & IN22)) | IN15)) & ((!(((((!(IN21)) & (!(IN2))) & IN1) & (!(IN20))) & IN22)) | IN12)) & ((!((((IN21 & (!(IN2))) & IN1) & (!(IN20))) & IN22)) | IN11)) & ((!(((((!(IN21)) & IN2) & IN1) & (!(IN20))) & IN22)) | IN9)) & ((!((((IN21 & IN2) & IN1) & (!(IN20))) & IN22)) | IN13)) & ((!(((((!(IN21)) & (!(IN2))) & (!(IN1))) & IN20) & IN22)) | IN27)) & ((!((((IN21 & (!(IN2))) & (!(IN1))) & IN20) & IN22)) | IN14)) & ((!(((((!(IN21)) & IN2) & (!(IN1))) & IN20) & IN22)) | IN31)) & ((!((((IN21 & IN2) & (!(IN1))) & IN20) & IN22)) | IN35)) & ((!(((((!(IN21)) & (!(IN2))) & IN1) & IN20) & IN22)) | IN36)) & ((!((((IN21 & (!(IN2))) & IN1) & IN20) & IN22)) | IN18)) & ((!(((((!(IN21)) & IN2) & IN1) & IN20) & IN22)) | IN19)) & ((!((((IN21 & IN2) & IN1) & IN20) & IN22)) | IN37)

*)

FUNCTION_BLOCK F_CollectInput
  VAR_IN_OUT
      Data : ARRAY[1..40] OF BOOL;
  END_VAR
  VAR_INPUT
      TICK  : BOOL := 0;
      IN1   : BOOL := 0;
      IN2   : BOOL := 0;
      IN3   : BOOL := 0;
      IN4   : BOOL := 0;
      IN5   : BOOL := 0;
      RESET : BOOL := FALSE;
  END_VAR
  VAR_OUTPUT
      Finished : BOOL;
  END_VAR
  VAR
      j    : USINT := 1;
      tock : BOOL  := 0;
  END_VAR
  IF NOT RESET AND tock = NOT TICK THEN
      Data[j]   := IN1;
      Data[j+1] := IN2;
      Data[j+2] := IN3;
      Data[j+3] := IN4;
      Data[j+4] := IN5;
      j := j + 5;
      tock := TICK;
  ELSE
      j := 1;
      tock := 0;
  END_IF;
  Finished := (j > 40);
END_FUNCTION_BLOCK

PROGRAM Boiler
  VAR
    Data  : ARRAY[1..40] OF BOOL;
    Ready : BOOL;
    CollectInput : F_CollectInput;
  END_VAR
  VAR
    TICK     AT %IX1.0 : BOOL;
    IN1      AT %IX0.3 : BOOL;
    IN2      AT %IX0.4 : BOOL;
    IN3      AT %IX0.5 : BOOL;
    IN4      AT %IX0.6 : BOOL;
    IN5      AT %IX0.7 : BOOL;
    OutReady AT %QX0.0 : BOOL := FALSE;
    FeedNext AT %QX0.1 : BOOL := FALSE;
    Out      AT %QX0.2 : BOOL;
  END_VAR
  CollectInput(TICK:=TICK, IN1:=IN1, IN2:=IN2, IN3:=IN3, IN4:=IN4, IN5:=IN5);
  Ready := CollectInput.Finished;
  FeedNext := 1;
  IF Ready THEN
    Out := (((((((((((((((((((((((((((((((((NOT (((((NOT Data[21]) AND (NOT Data[2])) AND (NOT Data[1])) AND (NOT Data[20])) AND (NOT Data[22]))) OR Data[3]) AND ((NOT ((((Data[21] AND (NOT Data[2])) AND (NOT Data[1])) AND (NOT Data[20])) AND (NOT Data[22]))) OR Data[24])) AND ((NOT (((((NOT Data[21]) AND Data[2]) AND (NOT Data[1])) AND (NOT Data[20])) AND (NOT Data[22]))) OR Data[23])) AND ((NOT ((((Data[21] AND Data[2]) AND (NOT Data[1])) AND (NOT Data[20])) AND (NOT Data[22]))) OR Data[25])) AND ((NOT (((((NOT Data[21]) AND (NOT Data[2])) AND Data[1]) AND (NOT Data[20])) AND (NOT Data[22]))) OR Data[28])) AND ((NOT ((((Data[21] AND (NOT Data[2])) AND Data[1]) AND (NOT Data[20])) AND (NOT Data[22]))) OR Data[6])) AND ((NOT (((((NOT Data[21]) AND Data[2]) AND Data[1]) AND (NOT Data[20])) AND (NOT Data[22]))) OR Data[4])) AND ((NOT ((((Data[21] AND Data[2]) AND Data[1]) AND (NOT Data[20])) AND (NOT Data[22]))) OR Data[26])) AND ((NOT (((((NOT Data[21]) AND (NOT Data[2])) AND (NOT Data[1])) AND Data[20]) AND (NOT Data[22]))) OR Data[29])) AND ((NOT ((((Data[21] AND (NOT Data[2])) AND (NOT Data[1])) AND Data[20]) AND (NOT Data[22]))) OR Data[30])) AND ((NOT (((((NOT Data[21]) AND Data[2]) AND (NOT Data[1])) AND Data[20]) AND (NOT Data[22]))) OR Data[7])) AND ((NOT ((((Data[21] AND Data[2]) AND (NOT Data[1])) AND Data[20]) AND (NOT Data[22]))) OR Data[8])) AND ((NOT (((((NOT Data[21]) AND (NOT Data[2])) AND Data[1]) AND Data[20]) AND (NOT Data[22]))) OR Data[34])) AND ((NOT ((((Data[21] AND (NOT Data[2])) AND Data[1]) AND Data[20]) AND (NOT Data[22]))) OR Data[5])) AND ((NOT (((((NOT Data[21]) AND Data[2]) AND Data[1]) AND Data[20]) AND (NOT Data[22]))) OR Data[16])) AND ((NOT ((((Data[21] AND Data[2]) AND Data[1]) AND Data[20]) AND (NOT Data[22]))) OR Data[17])) AND ((NOT (((((NOT Data[21]) AND (NOT Data[2])) AND (NOT Data[1])) AND (NOT Data[20])) AND Data[22])) OR Data[10])) AND ((NOT ((((Data[21] AND (NOT Data[2])) AND (NOT Data[1])) AND (NOT Data[20])) AND Data[22])) OR Data[32])) AND ((NOT (((((NOT Data[21]) AND Data[2]) AND (NOT Data[1])) AND (NOT Data[20])) AND Data[22])) OR Data[33])) AND ((NOT ((((Data[21] AND Data[2]) AND (NOT Data[1])) AND (NOT Data[20])) AND Data[22])) OR Data[15])) AND ((NOT (((((NOT Data[21]) AND (NOT Data[2])) AND Data[1]) AND (NOT Data[20])) AND Data[22])) OR Data[12])) AND ((NOT ((((Data[21] AND (NOT Data[2])) AND Data[1]) AND (NOT Data[20])) AND Data[22])) OR Data[11])) AND ((NOT (((((NOT Data[21]) AND Data[2]) AND Data[1]) AND (NOT Data[20])) AND Data[22])) OR Data[9])) AND ((NOT ((((Data[21] AND Data[2]) AND Data[1]) AND (NOT Data[20])) AND Data[22])) OR Data[13])) AND ((NOT (((((NOT Data[21]) AND (NOT Data[2])) AND (NOT Data[1])) AND Data[20]) AND Data[22])) OR Data[27])) AND ((NOT ((((Data[21] AND (NOT Data[2])) AND (NOT Data[1])) AND Data[20]) AND Data[22])) OR Data[14])) AND ((NOT (((((NOT Data[21]) AND Data[2]) AND (NOT Data[1])) AND Data[20]) AND Data[22])) OR Data[31])) AND ((NOT ((((Data[21] AND Data[2]) AND (NOT Data[1])) AND Data[20]) AND Data[22])) OR Data[35])) AND ((NOT (((((NOT Data[21]) AND (NOT Data[2])) AND Data[1]) AND Data[20]) AND Data[22])) OR Data[36])) AND ((NOT ((((Data[21] AND (NOT Data[2])) AND Data[1]) AND Data[20]) AND Data[22])) OR Data[18])) AND ((NOT (((((NOT Data[21]) AND Data[2]) AND Data[1]) AND Data[20]) AND Data[22])) OR Data[19])) AND ((NOT ((((Data[21] AND Data[2]) AND Data[1]) AND Data[20]) AND Data[22])) OR Data[37]));
    OutReady := 1;
    CollectInput(RESET:=TRUE);
  END_IF;
END_PROGRAM

CONFIGURATION Config0
  RESOURCE Res0 ON PLC
    TASK task0(INTERVAL := T#20ms,PRIORITY := 0);
    PROGRAM instance0 WITH task0 : Boiler;
  END_RESOURCE
END_CONFIGURATION

(* ---- 5-MUX_thees-ephah-coked.st ---- *)
(*
This code implements a shuffled multiplexer with 5 control bits.
The control bits are: Data[N3], Data[N23], Data[N22], Data[N2], Data[N5]
The input bits are: Data[N20], Data[N25], Data[N6], Data[N1], Data[N24], Data[N26], Data[N21], Data[N27], Data[N28], Data[N29], Data[N35], Data[N31], Data[N34], Data[N30], Data[N32], Data[N7], Data[N4], Data[N33], Data[N36], Data[N8], Data[N9], Data[N37], Data[N10], Data[N11], Data[N12], Data[N15], Data[N13], Data[N16], Data[N17], Data[N14], Data[N19], Data[N18]

The symbolic expression is:
((((((((((((((((((((((((((((((((!(((((!(IN3)) & (!(IN23))) & (!(IN22))) & (!(IN2))) & (!(IN5)))) | IN20) & ((!((((IN3 & (!(IN23))) & (!(IN22))) & (!(IN2))) & (!(IN5)))) | IN25)) & ((!(((((!(IN3)) & IN23) & (!(IN22))) & (!(IN2))) & (!(IN5)))) | IN6)) & ((!((((IN3 & IN23) & (!(IN22))) & (!(IN2))) & (!(IN5)))) | IN1)) & ((!(((((!(IN3)) & (!(IN23))) & IN22) & (!(IN2))) & (!(IN5)))) | IN24)) & ((!((((IN3 & (!(IN23))) & IN22) & (!(IN2))) & (!(IN5)))) | IN26)) & ((!(((((!(IN3)) & IN23) & IN22) & (!(IN2))) & (!(IN5)))) | IN21)) & ((!((((IN3 & IN23) & IN22) & (!(IN2))) & (!(IN5)))) | IN27)) & ((!(((((!(IN3)) & (!(IN23))) & (!(IN22))) & IN2) & (!(IN5)))) | IN28)) & ((!((((IN3 & (!(IN23))) & (!(IN22))) & IN2) & (!(IN5)))) | IN29)) & ((!(((((!(IN3)) & IN23) & (!(IN22))) & IN2) & (!(IN5)))) | IN35)) & ((!((((IN3 & IN23) & (!(IN22))) & IN2) & (!(IN5)))) | IN31)) & ((!(((((!(IN3)) & (!(IN23))) & IN22) & IN2) & (!(IN5)))) | IN34)) & ((!((((IN3 & (!(IN23))) & IN22) & IN2) & (!(IN5)))) | IN30)) & ((!(((((!(IN3)) & IN23) & IN22) & IN2) & (!(IN5)))) | IN32)) & ((!((((IN3 & IN23) & IN22) & IN2) & (!(IN5)))) | IN7)) & ((!(((((!(IN3)) & (!(IN23))) & (!(IN22))) & (!(IN2))) & IN5)) | IN4)) & ((!((((IN3 & (!(IN23))) & (!(IN22))) & (!(IN2))) & IN5)) | IN33)) & ((!(((((!(IN3)) & IN23) & (!(IN22))) & (!(IN2))) & IN5)) | IN36)) & ((!((((IN3 & IN23) & (!(IN22))) & (!(IN2))) & IN5)) | IN8)) & ((!(((((!(IN3)) & (!(IN23))) & IN22) & (!(IN2))) & IN5)) | IN9)) & ((!((((IN3 & (!(IN23))) & IN22) & (!(IN2))) & IN5)) | IN37)) & ((!(((((!(IN3)) & IN23) & IN22) & (!(IN2))) & IN5)) | IN10)) & ((!((((IN3 & IN23) & IN22) & (!(IN2))) & IN5)) | IN11)) & ((!(((((!(IN3)) & (!(IN23))) & (!(IN22))) & IN2) & IN5)) | IN12)) & ((!((((IN3 & (!(IN23))) & (!(IN22))) & IN2) & IN5)) | IN15)) & ((!(((((!(IN3)) & IN23) & (!(IN22))) & IN2) & IN5)) | IN13)) & ((!((((IN3 & IN23) & (!(IN22))) & IN2) & IN5)) | IN16)) & ((!(((((!(IN3)) & (!(IN23))) & IN22) & IN2) & IN5)) | IN17)) & ((!((((IN3 & (!(IN23))) & IN22) & IN2) & IN5)) | IN14)) & ((!(((((!(IN3)) & IN23) & IN22) & IN2) & IN5)) | IN19)) & ((!((((IN3 & IN23) & IN22) & IN2) & IN5)) | IN18)

*)

FUNCTION_BLOCK F_CollectInput
  VAR_IN_OUT
      Data : ARRAY[1..40] OF BOOL;
  END_VAR
  VAR_INPUT
      TICK  : BOOL := 0;
      IN1   : BOOL := 0;
      IN2   : BOOL := 0;
      IN3   : BOOL := 0;
      IN4   : BOOL := 0;
      IN5   : BOOL := 0;
      RESET : BOOL := FALSE;
  END_VAR
  VAR_OUTPUT
      Finished : BOOL;
  END_VAR
  VAR
      j    : USINT := 1;
      tock : BOOL  := 0;
  END_VAR
  IF NOT RESET AND tock = NOT TICK THEN
      Data[j]   := IN1;
      Data[j+1] := IN2;
      Data[j+2] := IN3;
      Data[j+3] := IN4;
      Data[j+4] := IN5;
      j := j + 5;
      tock := TICK;
  ELSE
      j := 1;
      tock := 0;
  END_IF;
  Finished := (j > 40);
END_FUNCTION_BLOCK

PROGRAM Boiler
  VAR
    Data  : ARRAY[1..40] OF BOOL;
    Ready : BOOL;
    CollectInput : F_CollectInput;
  END_VAR
  VAR
    TICK     AT %IX1.0 : BOOL;
    IN1      AT %IX0.3 : BOOL;
    IN2      AT %IX0.4 : BOOL;
    IN3      AT %IX0.5 : BOOL;
    IN4      AT %IX0.6 : BOOL;
    IN5      AT %IX0.7 : BOOL;
    OutReady AT %QX0.0 : BOOL := FALSE;
    FeedNext AT %QX0.1 : BOOL := FALSE;
    Out      AT %QX0.2 : BOOL;
  END_VAR
  CollectInput(TICK:=TICK, IN1:=IN1, IN2:=IN2, IN3:=IN3, IN4:=IN4, IN5:=IN5);
  Ready := CollectInput.Finished;
  FeedNext := 1;
  IF Ready THEN
    Out := (((((((((((((((((((((((((((((((((NOT (((((NOT Data[3]) AND (NOT Data[23])) AND (NOT Data[22])) AND (NOT Data[2])) AND (NOT Data[5]))) OR Data[20]) AND ((NOT ((((Data[3] AND (NOT Data[23])) AND (NOT Data[22])) AND (NOT Data[2])) AND (NOT Data[5]))) OR Data[25])) AND ((NOT (((((NOT Data[3]) AND Data[23]) AND (NOT Data[22])) AND (NOT Data[2])) AND (NOT Data[5]))) OR Data[6])) AND ((NOT ((((Data[3] AND Data[23]) AND (NOT Data[22])) AND (NOT Data[2])) AND (NOT Data[5]))) OR Data[1])) AND ((NOT (((((NOT Data[3]) AND (NOT Data[23])) AND Data[22]) AND (NOT Data[2])) AND (NOT Data[5]))) OR Data[24])) AND ((NOT ((((Data[3] AND (NOT Data[23])) AND Data[22]) AND (NOT Data[2])) AND (NOT Data[5]))) OR Data[26])) AND ((NOT (((((NOT Data[3]) AND Data[23]) AND Data[22]) AND (NOT Data[2])) AND (NOT Data[5]))) OR Data[21])) AND ((NOT ((((Data[3] AND Data[23]) AND Data[22]) AND (NOT Data[2])) AND (NOT Data[5]))) OR Data[27])) AND ((NOT (((((NOT Data[3]) AND (NOT Data[23])) AND (NOT Data[22])) AND Data[2]) AND (NOT Data[5]))) OR Data[28])) AND ((NOT ((((Data[3] AND (NOT Data[23])) AND (NOT Data[22])) AND Data[2]) AND (NOT Data[5]))) OR Data[29])) AND ((NOT (((((NOT Data[3]) AND Data[23]) AND (NOT Data[22])) AND Data[2]) AND (NOT Data[5]))) OR Data[35])) AND ((NOT ((((Data[3] AND Data[23]) AND (NOT Data[22])) AND Data[2]) AND (NOT Data[5]))) OR Data[31])) AND ((NOT (((((NOT Data[3]) AND (NOT Data[23])) AND Data[22]) AND Data[2]) AND (NOT Data[5]))) OR Data[34])) AND ((NOT ((((Data[3] AND (NOT Data[23])) AND Data[22]) AND Data[2]) AND (NOT Data[5]))) OR Data[30])) AND ((NOT (((((NOT Data[3]) AND Data[23]) AND Data[22]) AND Data[2]) AND (NOT Data[5]))) OR Data[32])) AND ((NOT ((((Data[3] AND Data[23]) AND Data[22]) AND Data[2]) AND (NOT Data[5]))) OR Data[7])) AND ((NOT (((((NOT Data[3]) AND (NOT Data[23])) AND (NOT Data[22])) AND (NOT Data[2])) AND Data[5])) OR Data[4])) AND ((NOT ((((Data[3] AND (NOT Data[23])) AND (NOT Data[22])) AND (NOT Data[2])) AND Data[5])) OR Data[33])) AND ((NOT (((((NOT Data[3]) AND Data[23]) AND (NOT Data[22])) AND (NOT Data[2])) AND Data[5])) OR Data[36])) AND ((NOT ((((Data[3] AND Data[23]) AND (NOT Data[22])) AND (NOT Data[2])) AND Data[5])) OR Data[8])) AND ((NOT (((((NOT Data[3]) AND (NOT Data[23])) AND Data[22]) AND (NOT Data[2])) AND Data[5])) OR Data[9])) AND ((NOT ((((Data[3] AND (NOT Data[23])) AND Data[22]) AND (NOT Data[2])) AND Data[5])) OR Data[37])) AND ((NOT (((((NOT Data[3]) AND Data[23]) AND Data[22]) AND (NOT Data[2])) AND Data[5])) OR Data[10])) AND ((NOT ((((Data[3] AND Data[23]) AND Data[22]) AND (NOT Data[2])) AND Data[5])) OR Data[11])) AND ((NOT (((((NOT Data[3]) AND (NOT Data[23])) AND (NOT Data[22])) AND Data[2]) AND Data[5])) OR Data[12])) AND ((NOT ((((Data[3] AND (NOT Data[23])) AND (NOT Data[22])) AND Data[2]) AND Data[5])) OR Data[15])) AND ((NOT (((((NOT Data[3]) AND Data[23]) AND (NOT Data[22])) AND Data[2]) AND Data[5])) OR Data[13])) AND ((NOT ((((Data[3] AND Data[23]) AND (NOT Data[22])) AND Data[2]) AND Data[5])) OR Data[16])) AND ((NOT (((((NOT Data[3]) AND (NOT Data[23])) AND Data[22]) AND Data[2]) AND Data[5])) OR Data[17])) AND ((NOT ((((Data[3] AND (NOT Data[23])) AND Data[22]) AND Data[2]) AND Data[5])) OR Data[14])) AND ((NOT (((((NOT Data[3]) AND Data[23]) AND Data[22]) AND Data[2]) AND Data[5])) OR Data[19])) AND ((NOT ((((Data[3] AND Data[23]) AND Data[22]) AND Data[2]) AND Data[5])) OR Data[18]));
    OutReady := 1;
    CollectInput(RESET:=TRUE);
  END_IF;
END_PROGRAM

CONFIGURATION Config0
  RESOURCE Res0 ON PLC
    TASK task0(INTERVAL := T#20ms,PRIORITY := 0);
    PROGRAM instance0 WITH task0 : Boiler;
  END_RESOURCE
END_CONFIGURATION

(* ---- 5-MUX_tight-duchy-saint.st ---- *)
(*
This code implements a shuffled multiplexer with 5 control bits.
The control bits are: Data[N21], Data[N20], Data[N2], Data[N1], Data[N3]
The input bits are: Data[N4], Data[N5], Data[N6], Data[N24], Data[N23], Data[N8], Data[N9], Data[N7], Data[N22], Data[N25], Data[N10], Data[N11], Data[N17], Data[N28], Data[N12], Data[N26], Data[N14], Data[N15], Data[N13], Data[N30], Data[N16], Data[N29], Data[N18], Data[N19], Data[N27], Data[N34], Data[N31], Data[N32], Data[N33], Data[N36], Data[N35], Data[N37]

The symbolic expression is:
((((((((((((((((((((((((((((((((!(((((!(IN21)) & (!(IN20))) & (!(IN2))) & (!(IN1))) & (!(IN3)))) | IN4) & ((!((((IN21 & (!(IN20))) & (!(IN2))) & (!(IN1))) & (!(IN3)))) | IN5)) & ((!(((((!(IN21)) & IN20) & (!(IN2))) & (!(IN1))) & (!(IN3)))) | IN6)) & ((!((((IN21 & IN20) & (!(IN2))) & (!(IN1))) & (!(IN3)))) | IN24)) & ((!(((((!(IN21)) & (!(IN20))) & IN2) & (!(IN1))) & (!(IN3)))) | IN23)) & ((!((((IN21 & (!(IN20))) & IN2) & (!(IN1))) & (!(IN3)))) | IN8)) & ((!(((((!(IN21)) & IN20) & IN2) & (!(IN1))) & (!(IN3)))) | IN9)) & ((!((((IN21 & IN20) & IN2) & (!(IN1))) & (!(IN3)))) | IN7)) & ((!(((((!(IN21)) & (!(IN20))) & (!(IN2))) & IN1) & (!(IN3)))) | IN22)) & ((!((((IN21 & (!(IN20))) & (!(IN2))) & IN1) & (!(IN3)))) | IN25)) & ((!(((((!(IN21)) & IN20) & (!(IN2))) & IN1) & (!(IN3)))) | IN10)) & ((!((((IN21 & IN20) & (!(IN2))) & IN1) & (!(IN3)))) | IN11)) & ((!(((((!(IN21)) & (!(IN20))) & IN2) & IN1) & (!(IN3)))) | IN17)) & ((!((((IN21 & (!(IN20))) & IN2) & IN1) & (!(IN3)))) | IN28)) & ((!(((((!(IN21)) & IN20) & IN2) & IN1) & (!(IN3)))) | IN12)) & ((!((((IN21 & IN20) & IN2) & IN1) & (!(IN3)))) | IN26)) & ((!(((((!(IN21)) & (!(IN20))) & (!(IN2))) & (!(IN1))) & IN3)) | IN14)) & ((!((((IN21 & (!(IN20))) & (!(IN2))) & (!(IN1))) & IN3)) | IN15)) & ((!(((((!(IN21)) & IN20) & (!(IN2))) & (!(IN1))) & IN3)) | IN13)) & ((!((((IN21 & IN20) & (!(IN2))) & (!(IN1))) & IN3)) | IN30)) & ((!(((((!(IN21)) & (!(IN20))) & IN2) & (!(IN1))) & IN3)) | IN16)) & ((!((((IN21 & (!(IN20))) & IN2) & (!(IN1))) & IN3)) | IN29)) & ((!(((((!(IN21)) & IN20) & IN2) & (!(IN1))) & IN3)) | IN18)) & ((!((((IN21 & IN20) & IN2) & (!(IN1))) & IN3)) | IN19)) & ((!(((((!(IN21)) & (!(IN20))) & (!(IN2))) & IN1) & IN3)) | IN27)) & ((!((((IN21 & (!(IN20))) & (!(IN2))) & IN1) & IN3)) | IN34)) & ((!(((((!(IN21)) & IN20) & (!(IN2))) & IN1) & IN3)) | IN31)) & ((!((((IN21 & IN20) & (!(IN2))) & IN1) & IN3)) | IN32)) & ((!(((((!(IN21)) & (!(IN20))) & IN2) & IN1) & IN3)) | IN33)) & ((!((((IN21 & (!(IN20))) & IN2) & IN1) & IN3)) | IN36)) & ((!(((((!(IN21)) & IN20) & IN2) & IN1) & IN3)) | IN35)) & ((!((((IN21 & IN20) & IN2) & IN1) & IN3)) | IN37)

*)

FUNCTION_BLOCK F_CollectInput
  VAR_IN_OUT
      Data : ARRAY[1..40] OF BOOL;
  END_VAR
  VAR_INPUT
      TICK  : BOOL := 0;
      IN1   : BOOL := 0;
      IN2   : BOOL := 0;
      IN3   : BOOL := 0;
      IN4   : BOOL := 0;
      IN5   : BOOL := 0;
      RESET : BOOL := FALSE;
  END_VAR
  VAR_OUTPUT
      Finished : BOOL;
  END_VAR
  VAR
      j    : USINT := 1;
      tock : BOOL  := 0;
  END_VAR
  IF NOT RESET AND tock = NOT TICK THEN
      Data[j]   := IN1;
      Data[j+1] := IN2;
      Data[j+2] := IN3;
      Data[j+3] := IN4;
      Data[j+4] := IN5;
      j := j + 5;
      tock := TICK;
  ELSE
      j := 1;
      tock := 0;
  END_IF;
  Finished := (j > 40);
END_FUNCTION_BLOCK

PROGRAM Boiler
  VAR
    Data  : ARRAY[1..40] OF BOOL;
    Ready : BOOL;
    CollectInput : F_CollectInput;
  END_VAR
  VAR
    TICK     AT %IX1.0 : BOOL;
    IN1      AT %IX0.3 : BOOL;
    IN2      AT %IX0.4 : BOOL;
    IN3      AT %IX0.5 : BOOL;
    IN4      AT %IX0.6 : BOOL;
    IN5      AT %IX0.7 : BOOL;
    OutReady AT %QX0.0 : BOOL := FALSE;
    FeedNext AT %QX0.1 : BOOL := FALSE;
    Out      AT %QX0.2 : BOOL;
  END_VAR
  CollectInput(TICK:=TICK, IN1:=IN1, IN2:=IN2, IN3:=IN3, IN4:=IN4, IN5:=IN5);
  Ready := CollectInput.Finished;
  FeedNext := 1;
  IF Ready THEN
    Out := (((((((((((((((((((((((((((((((((NOT (((((NOT Data[21]) AND (NOT Data[20])) AND (NOT Data[2])) AND (NOT Data[1])) AND (NOT Data[3]))) OR Data[4]) AND ((NOT ((((Data[21] AND (NOT Data[20])) AND (NOT Data[2])) AND (NOT Data[1])) AND (NOT Data[3]))) OR Data[5])) AND ((NOT (((((NOT Data[21]) AND Data[20]) AND (NOT Data[2])) AND (NOT Data[1])) AND (NOT Data[3]))) OR Data[6])) AND ((NOT ((((Data[21] AND Data[20]) AND (NOT Data[2])) AND (NOT Data[1])) AND (NOT Data[3]))) OR Data[24])) AND ((NOT (((((NOT Data[21]) AND (NOT Data[20])) AND Data[2]) AND (NOT Data[1])) AND (NOT Data[3]))) OR Data[23])) AND ((NOT ((((Data[21] AND (NOT Data[20])) AND Data[2]) AND (NOT Data[1])) AND (NOT Data[3]))) OR Data[8])) AND ((NOT (((((NOT Data[21]) AND Data[20]) AND Data[2]) AND (NOT Data[1])) AND (NOT Data[3]))) OR Data[9])) AND ((NOT ((((Data[21] AND Data[20]) AND Data[2]) AND (NOT Data[1])) AND (NOT Data[3]))) OR Data[7])) AND ((NOT (((((NOT Data[21]) AND (NOT Data[20])) AND (NOT Data[2])) AND Data[1]) AND (NOT Data[3]))) OR Data[22])) AND ((NOT ((((Data[21] AND (NOT Data[20])) AND (NOT Data[2])) AND Data[1]) AND (NOT Data[3]))) OR Data[25])) AND ((NOT (((((NOT Data[21]) AND Data[20]) AND (NOT Data[2])) AND Data[1]) AND (NOT Data[3]))) OR Data[10])) AND ((NOT ((((Data[21] AND Data[20]) AND (NOT Data[2])) AND Data[1]) AND (NOT Data[3]))) OR Data[11])) AND ((NOT (((((NOT Data[21]) AND (NOT Data[20])) AND Data[2]) AND Data[1]) AND (NOT Data[3]))) OR Data[17])) AND ((NOT ((((Data[21] AND (NOT Data[20])) AND Data[2]) AND Data[1]) AND (NOT Data[3]))) OR Data[28])) AND ((NOT (((((NOT Data[21]) AND Data[20]) AND Data[2]) AND Data[1]) AND (NOT Data[3]))) OR Data[12])) AND ((NOT ((((Data[21] AND Data[20]) AND Data[2]) AND Data[1]) AND (NOT Data[3]))) OR Data[26])) AND ((NOT (((((NOT Data[21]) AND (NOT Data[20])) AND (NOT Data[2])) AND (NOT Data[1])) AND Data[3])) OR Data[14])) AND ((NOT ((((Data[21] AND (NOT Data[20])) AND (NOT Data[2])) AND (NOT Data[1])) AND Data[3])) OR Data[15])) AND ((NOT (((((NOT Data[21]) AND Data[20]) AND (NOT Data[2])) AND (NOT Data[1])) AND Data[3])) OR Data[13])) AND ((NOT ((((Data[21] AND Data[20]) AND (NOT Data[2])) AND (NOT Data[1])) AND Data[3])) OR Data[30])) AND ((NOT (((((NOT Data[21]) AND (NOT Data[20])) AND Data[2]) AND (NOT Data[1])) AND Data[3])) OR Data[16])) AND ((NOT ((((Data[21] AND (NOT Data[20])) AND Data[2]) AND (NOT Data[1])) AND Data[3])) OR Data[29])) AND ((NOT (((((NOT Data[21]) AND Data[20]) AND Data[2]) AND (NOT Data[1])) AND Data[3])) OR Data[18])) AND ((NOT ((((Data[21] AND Data[20]) AND Data[2]) AND (NOT Data[1])) AND Data[3])) OR Data[19])) AND ((NOT (((((NOT Data[21]) AND (NOT Data[20])) AND (NOT Data[2])) AND Data[1]) AND Data[3])) OR Data[27])) AND ((NOT ((((Data[21] AND (NOT Data[20])) AND (NOT Data[2])) AND Data[1]) AND Data[3])) OR Data[34])) AND ((NOT (((((NOT Data[21]) AND Data[20]) AND (NOT Data[2])) AND Data[1]) AND Data[3])) OR Data[31])) AND ((NOT ((((Data[21] AND Data[20]) AND (NOT Data[2])) AND Data[1]) AND Data[3])) OR Data[32])) AND ((NOT (((((NOT Data[21]) AND (NOT Data[20])) AND Data[2]) AND Data[1]) AND Data[3])) OR Data[33])) AND ((NOT ((((Data[21] AND (NOT Data[20])) AND Data[2]) AND Data[1]) AND Data[3])) OR Data[36])) AND ((NOT (((((NOT Data[21]) AND Data[20]) AND Data[2]) AND Data[1]) AND Data[3])) OR Data[35])) AND ((NOT ((((Data[21] AND Data[20]) AND Data[2]) AND Data[1]) AND Data[3])) OR Data[37]));
    OutReady := 1;
    CollectInput(RESET:=TRUE);
  END_IF;
END_PROGRAM

CONFIGURATION Config0
  RESOURCE Res0 ON PLC
    TASK task0(INTERVAL := T#20ms,PRIORITY := 0);
    PROGRAM instance0 WITH task0 : Boiler;
  END_RESOURCE
END_CONFIGURATION

(* ---- 5-MUX_trade-sicko-parch.st ---- *)
(*
This code implements a shuffled multiplexer with 5 control bits.
The control bits are: Data[N20], Data[N2], Data[N1], Data[N21], Data[N22]
The input bits are: Data[N24], Data[N3], Data[N28], Data[N23], Data[N4], Data[N25], Data[N29], Data[N27], Data[N5], Data[N6], Data[N35], Data[N8], Data[N26], Data[N30], Data[N10], Data[N7], Data[N31], Data[N11], Data[N9], Data[N33], Data[N12], Data[N15], Data[N34], Data[N16], Data[N32], Data[N37], Data[N36], Data[N19], Data[N13], Data[N18], Data[N14], Data[N17]

The symbolic expression is:
((((((((((((((((((((((((((((((((!(((((!(IN20)) & (!(IN2))) & (!(IN1))) & (!(IN21))) & (!(IN22)))) | IN24) & ((!((((IN20 & (!(IN2))) & (!(IN1))) & (!(IN21))) & (!(IN22)))) | IN3)) & ((!(((((!(IN20)) & IN2) & (!(IN1))) & (!(IN21))) & (!(IN22)))) | IN28)) & ((!((((IN20 & IN2) & (!(IN1))) & (!(IN21))) & (!(IN22)))) | IN23)) & ((!(((((!(IN20)) & (!(IN2))) & IN1) & (!(IN21))) & (!(IN22)))) | IN4)) & ((!((((IN20 & (!(IN2))) & IN1) & (!(IN21))) & (!(IN22)))) | IN25)) & ((!(((((!(IN20)) & IN2) & IN1) & (!(IN21))) & (!(IN22)))) | IN29)) & ((!((((IN20 & IN2) & IN1) & (!(IN21))) & (!(IN22)))) | IN27)) & ((!(((((!(IN20)) & (!(IN2))) & (!(IN1))) & IN21) & (!(IN22)))) | IN5)) & ((!((((IN20 & (!(IN2))) & (!(IN1))) & IN21) & (!(IN22)))) | IN6)) & ((!(((((!(IN20)) & IN2) & (!(IN1))) & IN21) & (!(IN22)))) | IN35)) & ((!((((IN20 & IN2) & (!(IN1))) & IN21) & (!(IN22)))) | IN8)) & ((!(((((!(IN20)) & (!(IN2))) & IN1) & IN21) & (!(IN22)))) | IN26)) & ((!((((IN20 & (!(IN2))) & IN1) & IN21) & (!(IN22)))) | IN30)) & ((!(((((!(IN20)) & IN2) & IN1) & IN21) & (!(IN22)))) | IN10)) & ((!((((IN20 & IN2) & IN1) & IN21) & (!(IN22)))) | IN7)) & ((!(((((!(IN20)) & (!(IN2))) & (!(IN1))) & (!(IN21))) & IN22)) | IN31)) & ((!((((IN20 & (!(IN2))) & (!(IN1))) & (!(IN21))) & IN22)) | IN11)) & ((!(((((!(IN20)) & IN2) & (!(IN1))) & (!(IN21))) & IN22)) | IN9)) & ((!((((IN20 & IN2) & (!(IN1))) & (!(IN21))) & IN22)) | IN33)) & ((!(((((!(IN20)) & (!(IN2))) & IN1) & (!(IN21))) & IN22)) | IN12)) & ((!((((IN20 & (!(IN2))) & IN1) & (!(IN21))) & IN22)) | IN15)) & ((!(((((!(IN20)) & IN2) & IN1) & (!(IN21))) & IN22)) | IN34)) & ((!((((IN20 & IN2) & IN1) & (!(IN21))) & IN22)) | IN16)) & ((!(((((!(IN20)) & (!(IN2))) & (!(IN1))) & IN21) & IN22)) | IN32)) & ((!((((IN20 & (!(IN2))) & (!(IN1))) & IN21) & IN22)) | IN37)) & ((!(((((!(IN20)) & IN2) & (!(IN1))) & IN21) & IN22)) | IN36)) & ((!((((IN20 & IN2) & (!(IN1))) & IN21) & IN22)) | IN19)) & ((!(((((!(IN20)) & (!(IN2))) & IN1) & IN21) & IN22)) | IN13)) & ((!((((IN20 & (!(IN2))) & IN1) & IN21) & IN22)) | IN18)) & ((!(((((!(IN20)) & IN2) & IN1) & IN21) & IN22)) | IN14)) & ((!((((IN20 & IN2) & IN1) & IN21) & IN22)) | IN17)

*)

FUNCTION_BLOCK F_CollectInput
  VAR_IN_OUT
      Data : ARRAY[1..40] OF BOOL;
  END_VAR
  VAR_INPUT
      TICK  : BOOL := 0;
      IN1   : BOOL := 0;
      IN2   : BOOL := 0;
      IN3   : BOOL := 0;
      IN4   : BOOL := 0;
      IN5   : BOOL := 0;
      RESET : BOOL := FALSE;
  END_VAR
  VAR_OUTPUT
      Finished : BOOL;
  END_VAR
  VAR
      j    : USINT := 1;
      tock : BOOL  := 0;
  END_VAR
  IF NOT RESET AND tock = NOT TICK THEN
      Data[j]   := IN1;
      Data[j+1] := IN2;
      Data[j+2] := IN3;
      Data[j+3] := IN4;
      Data[j+4] := IN5;
      j := j + 5;
      tock := TICK;
  ELSE
      j := 1;
      tock := 0;
  END_IF;
  Finished := (j > 40);
END_FUNCTION_BLOCK

PROGRAM Boiler
  VAR
    Data  : ARRAY[1..40] OF BOOL;
    Ready : BOOL;
    CollectInput : F_CollectInput;
  END_VAR
  VAR
    TICK     AT %IX1.0 : BOOL;
    IN1      AT %IX0.3 : BOOL;
    IN2      AT %IX0.4 : BOOL;
    IN3      AT %IX0.5 : BOOL;
    IN4      AT %IX0.6 : BOOL;
    IN5      AT %IX0.7 : BOOL;
    OutReady AT %QX0.0 : BOOL := FALSE;
    FeedNext AT %QX0.1 : BOOL := FALSE;
    Out      AT %QX0.2 : BOOL;
  END_VAR
  CollectInput(TICK:=TICK, IN1:=IN1, IN2:=IN2, IN3:=IN3, IN4:=IN4, IN5:=IN5);
  Ready := CollectInput.Finished;
  FeedNext := 1;
  IF Ready THEN
    Out := (((((((((((((((((((((((((((((((((NOT (((((NOT Data[20]) AND (NOT Data[2])) AND (NOT Data[1])) AND (NOT Data[21])) AND (NOT Data[22]))) OR Data[24]) AND ((NOT ((((Data[20] AND (NOT Data[2])) AND (NOT Data[1])) AND (NOT Data[21])) AND (NOT Data[22]))) OR Data[3])) AND ((NOT (((((NOT Data[20]) AND Data[2]) AND (NOT Data[1])) AND (NOT Data[21])) AND (NOT Data[22]))) OR Data[28])) AND ((NOT ((((Data[20] AND Data[2]) AND (NOT Data[1])) AND (NOT Data[21])) AND (NOT Data[22]))) OR Data[23])) AND ((NOT (((((NOT Data[20]) AND (NOT Data[2])) AND Data[1]) AND (NOT Data[21])) AND (NOT Data[22]))) OR Data[4])) AND ((NOT ((((Data[20] AND (NOT Data[2])) AND Data[1]) AND (NOT Data[21])) AND (NOT Data[22]))) OR Data[25])) AND ((NOT (((((NOT Data[20]) AND Data[2]) AND Data[1]) AND (NOT Data[21])) AND (NOT Data[22]))) OR Data[29])) AND ((NOT ((((Data[20] AND Data[2]) AND Data[1]) AND (NOT Data[21])) AND (NOT Data[22]))) OR Data[27])) AND ((NOT (((((NOT Data[20]) AND (NOT Data[2])) AND (NOT Data[1])) AND Data[21]) AND (NOT Data[22]))) OR Data[5])) AND ((NOT ((((Data[20] AND (NOT Data[2])) AND (NOT Data[1])) AND Data[21]) AND (NOT Data[22]))) OR Data[6])) AND ((NOT (((((NOT Data[20]) AND Data[2]) AND (NOT Data[1])) AND Data[21]) AND (NOT Data[22]))) OR Data[35])) AND ((NOT ((((Data[20] AND Data[2]) AND (NOT Data[1])) AND Data[21]) AND (NOT Data[22]))) OR Data[8])) AND ((NOT (((((NOT Data[20]) AND (NOT Data[2])) AND Data[1]) AND Data[21]) AND (NOT Data[22]))) OR Data[26])) AND ((NOT ((((Data[20] AND (NOT Data[2])) AND Data[1]) AND Data[21]) AND (NOT Data[22]))) OR Data[30])) AND ((NOT (((((NOT Data[20]) AND Data[2]) AND Data[1]) AND Data[21]) AND (NOT Data[22]))) OR Data[10])) AND ((NOT ((((Data[20] AND Data[2]) AND Data[1]) AND Data[21]) AND (NOT Data[22]))) OR Data[7])) AND ((NOT (((((NOT Data[20]) AND (NOT Data[2])) AND (NOT Data[1])) AND (NOT Data[21])) AND Data[22])) OR Data[31])) AND ((NOT ((((Data[20] AND (NOT Data[2])) AND (NOT Data[1])) AND (NOT Data[21])) AND Data[22])) OR Data[11])) AND ((NOT (((((NOT Data[20]) AND Data[2]) AND (NOT Data[1])) AND (NOT Data[21])) AND Data[22])) OR Data[9])) AND ((NOT ((((Data[20] AND Data[2]) AND (NOT Data[1])) AND (NOT Data[21])) AND Data[22])) OR Data[33])) AND ((NOT (((((NOT Data[20]) AND (NOT Data[2])) AND Data[1]) AND (NOT Data[21])) AND Data[22])) OR Data[12])) AND ((NOT ((((Data[20] AND (NOT Data[2])) AND Data[1]) AND (NOT Data[21])) AND Data[22])) OR Data[15])) AND ((NOT (((((NOT Data[20]) AND Data[2]) AND Data[1]) AND (NOT Data[21])) AND Data[22])) OR Data[34])) AND ((NOT ((((Data[20] AND Data[2]) AND Data[1]) AND (NOT Data[21])) AND Data[22])) OR Data[16])) AND ((NOT (((((NOT Data[20]) AND (NOT Data[2])) AND (NOT Data[1])) AND Data[21]) AND Data[22])) OR Data[32])) AND ((NOT ((((Data[20] AND (NOT Data[2])) AND (NOT Data[1])) AND Data[21]) AND Data[22])) OR Data[37])) AND ((NOT (((((NOT Data[20]) AND Data[2]) AND (NOT Data[1])) AND Data[21]) AND Data[22])) OR Data[36])) AND ((NOT ((((Data[20] AND Data[2]) AND (NOT Data[1])) AND Data[21]) AND Data[22])) OR Data[19])) AND ((NOT (((((NOT Data[20]) AND (NOT Data[2])) AND Data[1]) AND Data[21]) AND Data[22])) OR Data[13])) AND ((NOT ((((Data[20] AND (NOT Data[2])) AND Data[1]) AND Data[21]) AND Data[22])) OR Data[18])) AND ((NOT (((((NOT Data[20]) AND Data[2]) AND Data[1]) AND Data[21]) AND Data[22])) OR Data[14])) AND ((NOT ((((Data[20] AND Data[2]) AND Data[1]) AND Data[21]) AND Data[22])) OR Data[17]));
    OutReady := 1;
    CollectInput(RESET:=TRUE);
  END_IF;
END_PROGRAM

CONFIGURATION Config0
  RESOURCE Res0 ON PLC
    TASK task0(INTERVAL := T#20ms,PRIORITY := 0);
    PROGRAM instance0 WITH task0 : Boiler;
  END_RESOURCE
END_CONFIGURATION

(* ---- 5-MUX_tubas-dived-baize.st ---- *)
(*
This code implements a shuffled multiplexer with 5 control bits.
The control bits are: Data[N21], Data[N20], Data[N24], Data[N2], Data[N22]
The input bits are: Data[N1], Data[N3], Data[N25], Data[N5], Data[N7], Data[N8], Data[N4], Data[N23], Data[N6], Data[N26], Data[N27], Data[N9], Data[N10], Data[N29], Data[N13], Data[N11], Data[N12], Data[N28], Data[N16], Data[N30], Data[N34], Data[N15], Data[N31], Data[N17], Data[N14], Data[N19], Data[N32], Data[N37], Data[N18], Data[N33], Data[N36], Data[N35]

The symbolic expression is:
((((((((((((((((((((((((((((((((!(((((!(IN21)) & (!(IN20))) & (!(IN24))) & (!(IN2))) & (!(IN22)))) | IN1) & ((!((((IN21 & (!(IN20))) & (!(IN24))) & (!(IN2))) & (!(IN22)))) | IN3)) & ((!(((((!(IN21)) & IN20) & (!(IN24))) & (!(IN2))) & (!(IN22)))) | IN25)) & ((!((((IN21 & IN20) & (!(IN24))) & (!(IN2))) & (!(IN22)))) | IN5)) & ((!(((((!(IN21)) & (!(IN20))) & IN24) & (!(IN2))) & (!(IN22)))) | IN7)) & ((!((((IN21 & (!(IN20))) & IN24) & (!(IN2))) & (!(IN22)))) | IN8)) & ((!(((((!(IN21)) & IN20) & IN24) & (!(IN2))) & (!(IN22)))) | IN4)) & ((!((((IN21 & IN20) & IN24) & (!(IN2))) & (!(IN22)))) | IN23)) & ((!(((((!(IN21)) & (!(IN20))) & (!(IN24))) & IN2) & (!(IN22)))) | IN6)) & ((!((((IN21 & (!(IN20))) & (!(IN24))) & IN2) & (!(IN22)))) | IN26)) & ((!(((((!(IN21)) & IN20) & (!(IN24))) & IN2) & (!(IN22)))) | IN27)) & ((!((((IN21 & IN20) & (!(IN24))) & IN2) & (!(IN22)))) | IN9)) & ((!(((((!(IN21)) & (!(IN20))) & IN24) & IN2) & (!(IN22)))) | IN10)) & ((!((((IN21 & (!(IN20))) & IN24) & IN2) & (!(IN22)))) | IN29)) & ((!(((((!(IN21)) & IN20) & IN24) & IN2) & (!(IN22)))) | IN13)) & ((!((((IN21 & IN20) & IN24) & IN2) & (!(IN22)))) | IN11)) & ((!(((((!(IN21)) & (!(IN20))) & (!(IN24))) & (!(IN2))) & IN22)) | IN12)) & ((!((((IN21 & (!(IN20))) & (!(IN24))) & (!(IN2))) & IN22)) | IN28)) & ((!(((((!(IN21)) & IN20) & (!(IN24))) & (!(IN2))) & IN22)) | IN16)) & ((!((((IN21 & IN20) & (!(IN24))) & (!(IN2))) & IN22)) | IN30)) & ((!(((((!(IN21)) & (!(IN20))) & IN24) & (!(IN2))) & IN22)) | IN34)) & ((!((((IN21 & (!(IN20))) & IN24) & (!(IN2))) & IN22)) | IN15)) & ((!(((((!(IN21)) & IN20) & IN24) & (!(IN2))) & IN22)) | IN31)) & ((!((((IN21 & IN20) & IN24) & (!(IN2))) & IN22)) | IN17)) & ((!(((((!(IN21)) & (!(IN20))) & (!(IN24))) & IN2) & IN22)) | IN14)) & ((!((((IN21 & (!(IN20))) & (!(IN24))) & IN2) & IN22)) | IN19)) & ((!(((((!(IN21)) & IN20) & (!(IN24))) & IN2) & IN22)) | IN32)) & ((!((((IN21 & IN20) & (!(IN24))) & IN2) & IN22)) | IN37)) & ((!(((((!(IN21)) & (!(IN20))) & IN24) & IN2) & IN22)) | IN18)) & ((!((((IN21 & (!(IN20))) & IN24) & IN2) & IN22)) | IN33)) & ((!(((((!(IN21)) & IN20) & IN24) & IN2) & IN22)) | IN36)) & ((!((((IN21 & IN20) & IN24) & IN2) & IN22)) | IN35)

*)

FUNCTION_BLOCK F_CollectInput
  VAR_IN_OUT
      Data : ARRAY[1..40] OF BOOL;
  END_VAR
  VAR_INPUT
      TICK  : BOOL := 0;
      IN1   : BOOL := 0;
      IN2   : BOOL := 0;
      IN3   : BOOL := 0;
      IN4   : BOOL := 0;
      IN5   : BOOL := 0;
      RESET : BOOL := FALSE;
  END_VAR
  VAR_OUTPUT
      Finished : BOOL;
  END_VAR
  VAR
      j    : USINT := 1;
      tock : BOOL  := 0;
  END_VAR
  IF NOT RESET AND tock = NOT TICK THEN
      Data[j]   := IN1;
      Data[j+1] := IN2;
      Data[j+2] := IN3;
      Data[j+3] := IN4;
      Data[j+4] := IN5;
      j := j + 5;
      tock := TICK;
  ELSE
      j := 1;
      tock := 0;
  END_IF;
  Finished := (j > 40);
END_FUNCTION_BLOCK

PROGRAM Boiler
  VAR
    Data  : ARRAY[1..40] OF BOOL;
    Ready : BOOL;
    CollectInput : F_CollectInput;
  END_VAR
  VAR
    TICK     AT %IX1.0 : BOOL;
    IN1      AT %IX0.3 : BOOL;
    IN2      AT %IX0.4 : BOOL;
    IN3      AT %IX0.5 : BOOL;
    IN4      AT %IX0.6 : BOOL;
    IN5      AT %IX0.7 : BOOL;
    OutReady AT %QX0.0 : BOOL := FALSE;
    FeedNext AT %QX0.1 : BOOL := FALSE;
    Out      AT %QX0.2 : BOOL;
  END_VAR
  CollectInput(TICK:=TICK, IN1:=IN1, IN2:=IN2, IN3:=IN3, IN4:=IN4, IN5:=IN5);
  Ready := CollectInput.Finished;
  FeedNext := 1;
  IF Ready THEN
    Out := (((((((((((((((((((((((((((((((((NOT (((((NOT Data[21]) AND (NOT Data[20])) AND (NOT Data[24])) AND (NOT Data[2])) AND (NOT Data[22]))) OR Data[1]) AND ((NOT ((((Data[21] AND (NOT Data[20])) AND (NOT Data[24])) AND (NOT Data[2])) AND (NOT Data[22]))) OR Data[3])) AND ((NOT (((((NOT Data[21]) AND Data[20]) AND (NOT Data[24])) AND (NOT Data[2])) AND (NOT Data[22]))) OR Data[25])) AND ((NOT ((((Data[21] AND Data[20]) AND (NOT Data[24])) AND (NOT Data[2])) AND (NOT Data[22]))) OR Data[5])) AND ((NOT (((((NOT Data[21]) AND (NOT Data[20])) AND Data[24]) AND (NOT Data[2])) AND (NOT Data[22]))) OR Data[7])) AND ((NOT ((((Data[21] AND (NOT Data[20])) AND Data[24]) AND (NOT Data[2])) AND (NOT Data[22]))) OR Data[8])) AND ((NOT (((((NOT Data[21]) AND Data[20]) AND Data[24]) AND (NOT Data[2])) AND (NOT Data[22]))) OR Data[4])) AND ((NOT ((((Data[21] AND Data[20]) AND Data[24]) AND (NOT Data[2])) AND (NOT Data[22]))) OR Data[23])) AND ((NOT (((((NOT Data[21]) AND (NOT Data[20])) AND (NOT Data[24])) AND Data[2]) AND (NOT Data[22]))) OR Data[6])) AND ((NOT ((((Data[21] AND (NOT Data[20])) AND (NOT Data[24])) AND Data[2]) AND (NOT Data[22]))) OR Data[26])) AND ((NOT (((((NOT Data[21]) AND Data[20]) AND (NOT Data[24])) AND Data[2]) AND (NOT Data[22]))) OR Data[27])) AND ((NOT ((((Data[21] AND Data[20]) AND (NOT Data[24])) AND Data[2]) AND (NOT Data[22]))) OR Data[9])) AND ((NOT (((((NOT Data[21]) AND (NOT Data[20])) AND Data[24]) AND Data[2]) AND (NOT Data[22]))) OR Data[10])) AND ((NOT ((((Data[21] AND (NOT Data[20])) AND Data[24]) AND Data[2]) AND (NOT Data[22]))) OR Data[29])) AND ((NOT (((((NOT Data[21]) AND Data[20]) AND Data[24]) AND Data[2]) AND (NOT Data[22]))) OR Data[13])) AND ((NOT ((((Data[21] AND Data[20]) AND Data[24]) AND Data[2]) AND (NOT Data[22]))) OR Data[11])) AND ((NOT (((((NOT Data[21]) AND (NOT Data[20])) AND (NOT Data[24])) AND (NOT Data[2])) AND Data[22])) OR Data[12])) AND ((NOT ((((Data[21] AND (NOT Data[20])) AND (NOT Data[24])) AND (NOT Data[2])) AND Data[22])) OR Data[28])) AND ((NOT (((((NOT Data[21]) AND Data[20]) AND (NOT Data[24])) AND (NOT Data[2])) AND Data[22])) OR Data[16])) AND ((NOT ((((Data[21] AND Data[20]) AND (NOT Data[24])) AND (NOT Data[2])) AND Data[22])) OR Data[30])) AND ((NOT (((((NOT Data[21]) AND (NOT Data[20])) AND Data[24]) AND (NOT Data[2])) AND Data[22])) OR Data[34])) AND ((NOT ((((Data[21] AND (NOT Data[20])) AND Data[24]) AND (NOT Data[2])) AND Data[22])) OR Data[15])) AND ((NOT (((((NOT Data[21]) AND Data[20]) AND Data[24]) AND (NOT Data[2])) AND Data[22])) OR Data[31])) AND ((NOT ((((Data[21] AND Data[20]) AND Data[24]) AND (NOT Data[2])) AND Data[22])) OR Data[17])) AND ((NOT (((((NOT Data[21]) AND (NOT Data[20])) AND (NOT Data[24])) AND Data[2]) AND Data[22])) OR Data[14])) AND ((NOT ((((Data[21] AND (NOT Data[20])) AND (NOT Data[24])) AND Data[2]) AND Data[22])) OR Data[19])) AND ((NOT (((((NOT Data[21]) AND Data[20]) AND (NOT Data[24])) AND Data[2]) AND Data[22])) OR Data[32])) AND ((NOT ((((Data[21] AND Data[20]) AND (NOT Data[24])) AND Data[2]) AND Data[22])) OR Data[37])) AND ((NOT (((((NOT Data[21]) AND (NOT Data[20])) AND Data[24]) AND Data[2]) AND Data[22])) OR Data[18])) AND ((NOT ((((Data[21] AND (NOT Data[20])) AND Data[24]) AND Data[2]) AND Data[22])) OR Data[33])) AND ((NOT (((((NOT Data[21]) AND Data[20]) AND Data[24]) AND Data[2]) AND Data[22])) OR Data[36])) AND ((NOT ((((Data[21] AND Data[20]) AND Data[24]) AND Data[2]) AND Data[22])) OR Data[35]));
    OutReady := 1;
    CollectInput(RESET:=TRUE);
  END_IF;
END_PROGRAM

CONFIGURATION Config0
  RESOURCE Res0 ON PLC
    TASK task0(INTERVAL := T#20ms,PRIORITY := 0);
    PROGRAM instance0 WITH task0 : Boiler;
  END_RESOURCE
END_CONFIGURATION

(* ---- 5-MUX_utero-smell-joule.st ---- *)
(*
This code implements a shuffled multiplexer with 5 control bits.
The control bits are: Data[N2], Data[N21], Data[N20], Data[N7], Data[N22]
The input bits are: Data[N1], Data[N23], Data[N25], Data[N5], Data[N29], Data[N28], Data[N3], Data[N26], Data[N6], Data[N13], Data[N10], Data[N4], Data[N24], Data[N8], Data[N30], Data[N14], Data[N11], Data[N18], Data[N9], Data[N19], Data[N27], Data[N12], Data[N32], Data[N34], Data[N17], Data[N16], Data[N15], Data[N31], Data[N36], Data[N33], Data[N35], Data[N37]

The symbolic expression is:
((((((((((((((((((((((((((((((((!(((((!(IN2)) & (!(IN21))) & (!(IN20))) & (!(IN7))) & (!(IN22)))) | IN1) & ((!((((IN2 & (!(IN21))) & (!(IN20))) & (!(IN7))) & (!(IN22)))) | IN23)) & ((!(((((!(IN2)) & IN21) & (!(IN20))) & (!(IN7))) & (!(IN22)))) | IN25)) & ((!((((IN2 & IN21) & (!(IN20))) & (!(IN7))) & (!(IN22)))) | IN5)) & ((!(((((!(IN2)) & (!(IN21))) & IN20) & (!(IN7))) & (!(IN22)))) | IN29)) & ((!((((IN2 & (!(IN21))) & IN20) & (!(IN7))) & (!(IN22)))) | IN28)) & ((!(((((!(IN2)) & IN21) & IN20) & (!(IN7))) & (!(IN22)))) | IN3)) & ((!((((IN2 & IN21) & IN20) & (!(IN7))) & (!(IN22)))) | IN26)) & ((!(((((!(IN2)) & (!(IN21))) & (!(IN20))) & IN7) & (!(IN22)))) | IN6)) & ((!((((IN2 & (!(IN21))) & (!(IN20))) & IN7) & (!(IN22)))) | IN13)) & ((!(((((!(IN2)) & IN21) & (!(IN20))) & IN7) & (!(IN22)))) | IN10)) & ((!((((IN2 & IN21) & (!(IN20))) & IN7) & (!(IN22)))) | IN4)) & ((!(((((!(IN2)) & (!(IN21))) & IN20) & IN7) & (!(IN22)))) | IN24)) & ((!((((IN2 & (!(IN21))) & IN20) & IN7) & (!(IN22)))) | IN8)) & ((!(((((!(IN2)) & IN21) & IN20) & IN7) & (!(IN22)))) | IN30)) & ((!((((IN2 & IN21) & IN20) & IN7) & (!(IN22)))) | IN14)) & ((!(((((!(IN2)) & (!(IN21))) & (!(IN20))) & (!(IN7))) & IN22)) | IN11)) & ((!((((IN2 & (!(IN21))) & (!(IN20))) & (!(IN7))) & IN22)) | IN18)) & ((!(((((!(IN2)) & IN21) & (!(IN20))) & (!(IN7))) & IN22)) | IN9)) & ((!((((IN2 & IN21) & (!(IN20))) & (!(IN7))) & IN22)) | IN19)) & ((!(((((!(IN2)) & (!(IN21))) & IN20) & (!(IN7))) & IN22)) | IN27)) & ((!((((IN2 & (!(IN21))) & IN20) & (!(IN7))) & IN22)) | IN12)) & ((!(((((!(IN2)) & IN21) & IN20) & (!(IN7))) & IN22)) | IN32)) & ((!((((IN2 & IN21) & IN20) & (!(IN7))) & IN22)) | IN34)) & ((!(((((!(IN2)) & (!(IN21))) & (!(IN20))) & IN7) & IN22)) | IN17)) & ((!((((IN2 & (!(IN21))) & (!(IN20))) & IN7) & IN22)) | IN16)) & ((!(((((!(IN2)) & IN21) & (!(IN20))) & IN7) & IN22)) | IN15)) & ((!((((IN2 & IN21) & (!(IN20))) & IN7) & IN22)) | IN31)) & ((!(((((!(IN2)) & (!(IN21))) & IN20) & IN7) & IN22)) | IN36)) & ((!((((IN2 & (!(IN21))) & IN20) & IN7) & IN22)) | IN33)) & ((!(((((!(IN2)) & IN21) & IN20) & IN7) & IN22)) | IN35)) & ((!((((IN2 & IN21) & IN20) & IN7) & IN22)) | IN37)

*)

FUNCTION_BLOCK F_CollectInput
  VAR_IN_OUT
      Data : ARRAY[1..40] OF BOOL;
  END_VAR
  VAR_INPUT
      TICK  : BOOL := 0;
      IN1   : BOOL := 0;
      IN2   : BOOL := 0;
      IN3   : BOOL := 0;
      IN4   : BOOL := 0;
      IN5   : BOOL := 0;
      RESET : BOOL := FALSE;
  END_VAR
  VAR_OUTPUT
      Finished : BOOL;
  END_VAR
  VAR
      j    : USINT := 1;
      tock : BOOL  := 0;
  END_VAR
  IF NOT RESET AND tock = NOT TICK THEN
      Data[j]   := IN1;
      Data[j+1] := IN2;
      Data[j+2] := IN3;
      Data[j+3] := IN4;
      Data[j+4] := IN5;
      j := j + 5;
      tock := TICK;
  ELSE
      j := 1;
      tock := 0;
  END_IF;
  Finished := (j > 40);
END_FUNCTION_BLOCK

PROGRAM Boiler
  VAR
    Data  : ARRAY[1..40] OF BOOL;
    Ready : BOOL;
    CollectInput : F_CollectInput;
  END_VAR
  VAR
    TICK     AT %IX1.0 : BOOL;
    IN1      AT %IX0.3 : BOOL;
    IN2      AT %IX0.4 : BOOL;
    IN3      AT %IX0.5 : BOOL;
    IN4      AT %IX0.6 : BOOL;
    IN5      AT %IX0.7 : BOOL;
    OutReady AT %QX0.0 : BOOL := FALSE;
    FeedNext AT %QX0.1 : BOOL := FALSE;
    Out      AT %QX0.2 : BOOL;
  END_VAR
  CollectInput(TICK:=TICK, IN1:=IN1, IN2:=IN2, IN3:=IN3, IN4:=IN4, IN5:=IN5);
  Ready := CollectInput.Finished;
  FeedNext := 1;
  IF Ready THEN
    Out := (((((((((((((((((((((((((((((((((NOT (((((NOT Data[2]) AND (NOT Data[21])) AND (NOT Data[20])) AND (NOT Data[7])) AND (NOT Data[22]))) OR Data[1]) AND ((NOT ((((Data[2] AND (NOT Data[21])) AND (NOT Data[20])) AND (NOT Data[7])) AND (NOT Data[22]))) OR Data[23])) AND ((NOT (((((NOT Data[2]) AND Data[21]) AND (NOT Data[20])) AND (NOT Data[7])) AND (NOT Data[22]))) OR Data[25])) AND ((NOT ((((Data[2] AND Data[21]) AND (NOT Data[20])) AND (NOT Data[7])) AND (NOT Data[22]))) OR Data[5])) AND ((NOT (((((NOT Data[2]) AND (NOT Data[21])) AND Data[20]) AND (NOT Data[7])) AND (NOT Data[22]))) OR Data[29])) AND ((NOT ((((Data[2] AND (NOT Data[21])) AND Data[20]) AND (NOT Data[7])) AND (NOT Data[22]))) OR Data[28])) AND ((NOT (((((NOT Data[2]) AND Data[21]) AND Data[20]) AND (NOT Data[7])) AND (NOT Data[22]))) OR Data[3])) AND ((NOT ((((Data[2] AND Data[21]) AND Data[20]) AND (NOT Data[7])) AND (NOT Data[22]))) OR Data[26])) AND ((NOT (((((NOT Data[2]) AND (NOT Data[21])) AND (NOT Data[20])) AND Data[7]) AND (NOT Data[22]))) OR Data[6])) AND ((NOT ((((Data[2] AND (NOT Data[21])) AND (NOT Data[20])) AND Data[7]) AND (NOT Data[22]))) OR Data[13])) AND ((NOT (((((NOT Data[2]) AND Data[21]) AND (NOT Data[20])) AND Data[7]) AND (NOT Data[22]))) OR Data[10])) AND ((NOT ((((Data[2] AND Data[21]) AND (NOT Data[20])) AND Data[7]) AND (NOT Data[22]))) OR Data[4])) AND ((NOT (((((NOT Data[2]) AND (NOT Data[21])) AND Data[20]) AND Data[7]) AND (NOT Data[22]))) OR Data[24])) AND ((NOT ((((Data[2] AND (NOT Data[21])) AND Data[20]) AND Data[7]) AND (NOT Data[22]))) OR Data[8])) AND ((NOT (((((NOT Data[2]) AND Data[21]) AND Data[20]) AND Data[7]) AND (NOT Data[22]))) OR Data[30])) AND ((NOT ((((Data[2] AND Data[21]) AND Data[20]) AND Data[7]) AND (NOT Data[22]))) OR Data[14])) AND ((NOT (((((NOT Data[2]) AND (NOT Data[21])) AND (NOT Data[20])) AND (NOT Data[7])) AND Data[22])) OR Data[11])) AND ((NOT ((((Data[2] AND (NOT Data[21])) AND (NOT Data[20])) AND (NOT Data[7])) AND Data[22])) OR Data[18])) AND ((NOT (((((NOT Data[2]) AND Data[21]) AND (NOT Data[20])) AND (NOT Data[7])) AND Data[22])) OR Data[9])) AND ((NOT ((((Data[2] AND Data[21]) AND (NOT Data[20])) AND (NOT Data[7])) AND Data[22])) OR Data[19])) AND ((NOT (((((NOT Data[2]) AND (NOT Data[21])) AND Data[20]) AND (NOT Data[7])) AND Data[22])) OR Data[27])) AND ((NOT ((((Data[2] AND (NOT Data[21])) AND Data[20]) AND (NOT Data[7])) AND Data[22])) OR Data[12])) AND ((NOT (((((NOT Data[2]) AND Data[21]) AND Data[20]) AND (NOT Data[7])) AND Data[22])) OR Data[32])) AND ((NOT ((((Data[2] AND Data[21]) AND Data[20]) AND (NOT Data[7])) AND Data[22])) OR Data[34])) AND ((NOT (((((NOT Data[2]) AND (NOT Data[21])) AND (NOT Data[20])) AND Data[7]) AND Data[22])) OR Data[17])) AND ((NOT ((((Data[2] AND (NOT Data[21])) AND (NOT Data[20])) AND Data[7]) AND Data[22])) OR Data[16])) AND ((NOT (((((NOT Data[2]) AND Data[21]) AND (NOT Data[20])) AND Data[7]) AND Data[22])) OR Data[15])) AND ((NOT ((((Data[2] AND Data[21]) AND (NOT Data[20])) AND Data[7]) AND Data[22])) OR Data[31])) AND ((NOT (((((NOT Data[2]) AND (NOT Data[21])) AND Data[20]) AND Data[7]) AND Data[22])) OR Data[36])) AND ((NOT ((((Data[2] AND (NOT Data[21])) AND Data[20]) AND Data[7]) AND Data[22])) OR Data[33])) AND ((NOT (((((NOT Data[2]) AND Data[21]) AND Data[20]) AND Data[7]) AND Data[22])) OR Data[35])) AND ((NOT ((((Data[2] AND Data[21]) AND Data[20]) AND Data[7]) AND Data[22])) OR Data[37]));
    OutReady := 1;
    CollectInput(RESET:=TRUE);
  END_IF;
END_PROGRAM

CONFIGURATION Config0
  RESOURCE Res0 ON PLC
    TASK task0(INTERVAL := T#20ms,PRIORITY := 0);
    PROGRAM instance0 WITH task0 : Boiler;
  END_RESOURCE
END_CONFIGURATION
